FUNCTION_BLOCK "Auto_Test"   // FB1, SCL
{ S7_Optimized_Access := 'TRUE' }
VERSION : 0.1
// stored: AutoNumber true, IsIECCheckEnabled false, IsRetainMemResEnabled false, MemoryReserve 100, SetENOAutomatically false, UDAEnableTagReadback false
   VAR_INPUT
      Sys_No : UInt;
      Automatic : Bool;
      Manual : Bool;
      Level : UInt;
      Error : Bool;
      Start : Bool;
      Pause : Bool;
      Stop : Bool;
      "Pallet Type" : Char;
      "Tower 1 Pallet Alignment" : Char;
      "Tower 2 Pallet Alignment" : Char;
      "Extractor Pallet Alignment" : Char;
      Pallet_Allignment : Char;
      Tower : UInt;
      Transfer_From_To : Byte;
      "From level" : Byte;
      "To level" : Byte;
      "Testing Time" : UInt;
      "Numer of cycles" : Byte;
   END_VAR
   VAR_OUTPUT
      Running : Bool;
      Time_Runnng : Time;
      Start_Time { ExternalAccessible := 'False'; ExternalVisible := 'False'; ExternalWritable := 'False'} : String;
      Stop_Time { ExternalAccessible := 'False'; ExternalVisible := 'False'; ExternalWritable := 'False'} : String;
      Duration : Time;
   END_VAR
   VAR_IN_OUT
      "Order Table_1" : "OrderTable_UDT";
      Step_Table_0 : "OrderTable_UDT";
      System_OrderSent : Bool;
      Total_Duration : Time;
   END_VAR
   VAR
      State : Int;
      R_Start { S7_SetPoint := 'True'} : R_TRIG;
      T_Delay { S7_SetPoint := 'True'} : TON_TIME;
      Time_Delay : Time := T#0ms;
      Send_VTD_Order : Bool;
      Send_CNV_Order : Bool;
      R_TRIG_Instance { S7_SetPoint := 'True'} : R_TRIG;
      T_Running { S7_SetPoint := 'True'} : TON_TIME;
      F_TRIG { S7_SetPoint := 'True'} : F_TRIG;
      R_TRIG { S7_SetPoint := 'True'} : R_TRIG;
      Error_Code : Int;
      test : Bool;
      N_Cycles : UInt;
      Testing_Time : Time;
      R_Manual_Mode { S7_SetPoint := 'True'} : R_TRIG;
   END_VAR
   VAR_TEMP
      Busy : Bool;
   END_VAR
   VAR CONSTANT
      VTD_DEVICE : String := 'VTD';
      PALLET_INOUT_DEVICE : String := 'Pallet In Out';
      SHUTTLE_INOUT_DEVICE : String := 'Shuttle In Out';
      RUNNING_STATUS : String := 'Running';
      COMPLETED_STATUS : String := 'Completed';
   END_VAR
BEGIN
   #R_Start(CLK:=#Start);

   IF #Stop THEN
       #State := 0;
   END_IF;

   IF #Error THEN
       #State := 400;
   END_IF;

   #R_Manual_Mode(CLK:=#Automatic AND NOT #Error AND #Manual AND NOT #Running);

   IF #R_Manual_Mode.Q THEN
       #State := 500;
   ELSIF #Automatic AND NOT #Error AND NOT #Manual AND #State = 500 THEN
       #State := 0;
   END_IF;

   IF #State > 10 AND #State < 400 THEN
       #Running := TRUE;
   END_IF;

   //Time running
   #R_TRIG(CLK:=#Running);
   IF #R_TRIG.Q THEN
       #Start_Time := "Time".CurrentLocalTime;
       #Stop_Time := '';
   END_IF;
   #F_TRIG(CLK:=#Running);
   IF #F_TRIG.Q THEN
       #Duration := #T_Running.ET;
       #Total_Duration := #Duration + #Total_Duration;
       #Stop_Time := "Time".CurrentLocalTime;
   END_IF;
   #T_Running(IN:=#Running AND NOT #Pause,
                         PT:=t#24h);

   #Time_Runnng := #T_Running.ET;

   #Testing_Time := UINT_TO_TIME(#"Testing Time") * 60000;

   #Error_Code := WRIT_DBL(REQ := #test, SRCBLK := "Auto_Test_DB",BUSY=>#Busy, DSTBLK => "Auto_Test_DB");

   CASE #State OF
       0://Initialization
           #Running := false;
           #State := #State + 10;

       10://Idle
           IF #R_Start.Q AND #Automatic AND NOT #Error AND #"Pallet Type" <> '' AND #"From level" > 0 AND #"To level" > 0  THEN
               #N_Cycles := 0;
               #State := #State + 10;
           END_IF;

       20: //VTD TO START LEVEL
           IF "Control_DB".VTD_Sys[#Sys_No].Current_Level <> #"From level" THEN
               "VTD_Order_FC"(i_Sys := #Sys_No,
                              Level := #"From level",
                              StepTable_0 := #Step_Table_0);
               #R_TRIG_Instance(CLK := TRUE,
                                Q => #System_OrderSent);
               #T_Delay(IN := TRUE,
                        PT := #Time_Delay);
               IF #"Order Table_1".Status = #RUNNING_STATUS AND #T_Delay.Q THEN
                   #R_TRIG_Instance(CLK := FALSE,
                                    Q => #System_OrderSent);
                   #T_Delay(IN := FALSE,
                            PT := T#0ms);
                   #State := #State + 10;
               END_IF;
           ELSE
               #State := #State + 20;
           END_IF;

       30: //ACK VTD
           //Wait to complete and send ack
           IF #"Order Table_1".Status = #COMPLETED_STATUS AND NOT #Pause THEN
               "Control_DB".WCS_OPC_Control[#Sys_No].Movement_Request_Complete_Ack := TRUE;
               #State := #State + 10;
           END_IF;

       40: //CNV1
           "CNV_Order_FC"(i_Sys := #Sys_No,
                          Level := "Control_DB".VTD_Sys[#Sys_No].Current_Level,
                          Tower := 1,
                          Transfer_From_To := 2,
                          Pallet_Type := #"Pallet Type",
                          Pallet_Allignment := #"Tower 1 Pallet Alignment",
                          Device:=#PALLET_INOUT_DEVICE,
                          Task_Type:=4,
                          StepTable_0 := #Step_Table_0);
           #System_OrderSent := TRUE;
           #State := #State + 10;

       50: //RESET ACK
           IF #"Order Table_1".Status = #RUNNING_STATUS THEN
               "Control_DB".WCS_OPC_Control[#Sys_No].Movement_Request_Complete_Ack := FALSE;
               #R_TRIG_Instance(CLK := FALSE,
                                Q => #System_OrderSent);
               #State := #State + 10;
           END_IF;

       60: //ACK CNV1
           //Wait to complete and send ack
           IF #"Order Table_1".Status = #COMPLETED_STATUS AND NOT #Pause THEN
               "Control_DB".WCS_OPC_Control[#Sys_No].Movement_Request_Complete_Ack := TRUE;
               #State := #State + 10;
           END_IF;

       70: //ECVN TO TOWER 1
           "CNV_Order_FC"(i_Sys := #Sys_No,
                          Level := "Control_DB".VTD_Sys[#Sys_No].Current_Level,
                          Tower := 1,
                          Transfer_From_To := 1,
                          Pallet_Type := #"Pallet Type",
                          Pallet_Allignment := #"Extractor Pallet Alignment",
                          Device:=#PALLET_INOUT_DEVICE,
                          Task_Type:=4,
                          StepTable_0 := #Step_Table_0);
           #System_OrderSent := TRUE;
           #State := #State + 10;

       80: //RESET ACK
           IF #"Order Table_1".Status = #RUNNING_STATUS THEN
               "Control_DB".WCS_OPC_Control[#Sys_No].Movement_Request_Complete_Ack := FALSE;
               #State := #State + 10;
           END_IF;

       90: //ACK ECVN
           //Wait to complete and send ack
           IF #"Order Table_1".Status = #COMPLETED_STATUS AND NOT #Pause THEN
               "Control_DB".WCS_OPC_Control[#Sys_No].Movement_Request_Complete_Ack := TRUE;
               #State := #State + 10;
           END_IF;

       100: //VTD FROM START LEVEL TO FINAL LEVEL
           IF "Control_DB".VTD_Sys[#Sys_No].Current_Level < #"To level" THEN
               "VTD_Order_FC"(i_Sys := #Sys_No,
                              Level := "Control_DB".VTD_Sys[#Sys_No].Current_Level + 1,
                              StepTable_0 := #Step_Table_0);
               #System_OrderSent := TRUE;
               #State := #State + 10;
           ELSE
               #State := 130;
           END_IF;

       110: //RESET ACK
           IF #"Order Table_1".Status = #RUNNING_STATUS THEN
               "Control_DB".WCS_OPC_Control[#Sys_No].Movement_Request_Complete_Ack := FALSE;
               #State := #State + 10;
           END_IF;


       120: //ACK VTD
           //Wait to complete and send ack
           IF #"Order Table_1".Status = #COMPLETED_STATUS AND NOT #Pause THEN
               "Control_DB".WCS_OPC_Control[#Sys_No].Movement_Request_Complete_Ack := TRUE;
               #State := 40;
           END_IF;

       130: //VTD TO START LEVEL---------------------------------------------------------------------------------------------------
           "VTD_Order_FC"(i_Sys := #Sys_No,
                          Level := #"From level",
                          StepTable_0 := #Step_Table_0);
           #System_OrderSent := TRUE;
           #State := #State + 10;

       140: //RESET ACK
           IF #"Order Table_1".Status = #RUNNING_STATUS THEN
               "Control_DB".WCS_OPC_Control[#Sys_No].Movement_Request_Complete_Ack := FALSE;
               #State := #State + 10;
           END_IF;

       150: //ACK VTD START LEVEL
           //Wait to complete and send ack
           IF #Sys_No <= 3 THEN
               IF #"Order Table_1".Status = #COMPLETED_STATUS AND NOT #Pause THEN
                   "Control_DB".WCS_OPC_Control[#Sys_No].Movement_Request_Complete_Ack := TRUE;
                   #State := #State + 10;
               END_IF;
           ELSE
               IF #"Order Table_1".Status = #COMPLETED_STATUS AND NOT #Pause THEN
                   "Control_DB".WCS_OPC_Control[#Sys_No].Movement_Request_Complete_Ack := TRUE;
                   #State := 40; //TEST JUST CONV 1 FOR SYSTEM 4 AND 5
               END_IF;
           END_IF;

       160: //CNV2
           "CNV_Order_FC"(i_Sys := #Sys_No,
                          Level := "Control_DB".VTD_Sys[#Sys_No].Current_Level,
                          Tower := 2,
                          Transfer_From_To := 2,
                          Pallet_Type := #"Pallet Type",
                          Pallet_Allignment := #"Tower 2 Pallet Alignment",
                          Device:=#PALLET_INOUT_DEVICE,
                          Task_Type:=4,
                          StepTable_0 := #Step_Table_0);
           #System_OrderSent := TRUE;
           #State := #State + 10;

       170: //RESET ACK
           IF #"Order Table_1".Status = #RUNNING_STATUS THEN
               "Control_DB".WCS_OPC_Control[#Sys_No].Movement_Request_Complete_Ack := FALSE;
               #State := #State + 10;
           END_IF;

       180: //ACK CNV2
           //Wait to complete and send ack
           IF #"Order Table_1".Status = #COMPLETED_STATUS AND NOT #Pause THEN
               "Control_DB".WCS_OPC_Control[#Sys_No].Movement_Request_Complete_Ack := TRUE;
               #State := #State + 10;
           END_IF;

       190: //ECVN TO TOWER 2
           "CNV_Order_FC"(i_Sys := #Sys_No,
                          Level := "Control_DB".VTD_Sys[#Sys_No].Current_Level,
                          Tower := 2,
                          Transfer_From_To := 1,
                          Pallet_Type := #"Pallet Type",
                          Pallet_Allignment := #"Extractor Pallet Alignment",
                          Device:=#PALLET_INOUT_DEVICE,
                          Task_Type:=4,
                          StepTable_0 := #Step_Table_0);
           #System_OrderSent := TRUE;
           #State := #State + 10;

       200: //RESET ACK
           IF #"Order Table_1".Status = #RUNNING_STATUS THEN
               "Control_DB".WCS_OPC_Control[#Sys_No].Movement_Request_Complete_Ack := FALSE;
               #State := #State + 10;
           END_IF;

       210: //ACK ECVN TO TOWER 2
           //Wait to complete and send ack
           IF #"Order Table_1".Status = #COMPLETED_STATUS AND NOT #Pause THEN
               "Control_DB".WCS_OPC_Control[#Sys_No].Movement_Request_Complete_Ack := TRUE;
               #State := #State + 10;
           END_IF;

       220: //VTD 
           IF "Control_DB".VTD_Sys[#Sys_No].Current_Level < #"To level" THEN
               "VTD_Order_FC"(i_Sys := #Sys_No,
                              Level := "Control_DB".VTD_Sys[#Sys_No].Current_Level + 1,
                              StepTable_0 := #Step_Table_0);
               #System_OrderSent := TRUE;
               #State := #State + 10;
           ELSIF (
               (#"Numer of cycles" = 0 OR #N_Cycles < #"Numer of cycles")
               AND
               (#Testing_Time = T#0M OR #Time_Runnng < #Testing_Time)
               ) THEN
               #State := 250;//CONTINUE
           ELSE
               #State := 260;//FINISH
           END_IF;

       230: //RESET ACK
           IF #"Order Table_1".Status = #RUNNING_STATUS THEN
               "Control_DB".WCS_OPC_Control[#Sys_No].Movement_Request_Complete_Ack := FALSE;
               #State := #State + 10;
           END_IF;

       240: //ACK VTD
           //Wait to complete and send ack
           IF #"Order Table_1".Status = #COMPLETED_STATUS AND NOT #Pause THEN
               "Control_DB".WCS_OPC_Control[#Sys_No].Movement_Request_Complete_Ack := TRUE;
               #State := 160;
           END_IF;

       250: //ACK VTD AND START ANOTHER CYCLE
           //Wait to complete and send ack
           IF #"Order Table_1".Status = #COMPLETED_STATUS AND NOT #Pause THEN
               "Control_DB".WCS_OPC_Control[#Sys_No].Movement_Request_Complete_Ack := TRUE;
               #N_Cycles := #N_Cycles + 1;
               #State := 20;
           END_IF;

       260: //ACK VTD AND FINISH
           //Wait to complete and send ack
           IF #"Order Table_1".Status = #COMPLETED_STATUS AND NOT #Pause THEN
               "Control_DB".WCS_OPC_Control[#Sys_No].Movement_Request_Complete_Ack := TRUE;
               #State := 0;
           END_IF;

       400: //ERROR
           #Running := false;
           IF "Reset_All" OR
               ("Screen_DB_1".Reset_All[1] AND
                ("HMI_Box_Connected_1" = 1) OR ("HMI_Box_Connected_1" = 2) OR ("HMI_Box_Connected_1" = 3) OR ("HMI_Box_Connected_1" = 4) OR ("HMI_Box_Connected_1" = 5) OR
                ("HMI_Box_Connected_1" = 11 AND "KEY REMOTE/LOCAL L1 - CH1(1)") OR
                ("HMI_Box_Connected_1" = 12 AND "KEY REMOTE/LOCAL L2 - CH1(1)") OR
                ("HMI_Box_Connected_1" = 13 AND "KEY REMOTE/LOCAL L3 - CH1(1)") OR
                ("HMI_Box_Connected_1" = 14 AND "KEY REMOTE/LOCAL L4 - CH1(1)") OR
                ("HMI_Box_Connected_1" = 15 AND "KEY REMOTE/LOCAL L5 - CH1(1)") OR
                ("HMI_Box_Connected_1" = 16 AND "KEY REMOTE/LOCAL L6 - CH1(1)") OR
                ("HMI_Box_Connected_1" = 17 AND "KEY REMOTE/LOCAL L7 - CH1(1)") OR
                ("HMI_Box_Connected_1" = 18 AND "KEY REMOTE/LOCAL L8 - CH1(1)") OR
                ("HMI_Box_Connected_1" = 21 AND "KEY REMOTE/LOCAL L1 - CH1(2)") OR
                ("HMI_Box_Connected_1" = 22 AND "KEY REMOTE/LOCAL L2 - CH1(2)") OR
                ("HMI_Box_Connected_1" = 23 AND "KEY REMOTE/LOCAL L3 - CH1(2)") OR
                ("HMI_Box_Connected_1" = 24 AND "KEY REMOTE/LOCAL L4 - CH1(2)") OR
                ("HMI_Box_Connected_1" = 25 AND "KEY REMOTE/LOCAL L5 - CH1(2)") OR
                ("HMI_Box_Connected_1" = 26 AND "KEY REMOTE/LOCAL L6 - CH1(2)") OR
                ("HMI_Box_Connected_1" = 27 AND "KEY REMOTE/LOCAL L7 - CH1(2)") OR
                ("HMI_Box_Connected_1" = 28 AND "KEY REMOTE/LOCAL L8 - CH1(2)") OR
                ("HMI_Box_Connected_1" = 31 AND "KEY REMOTE/LOCAL L1 - CH1(3)") OR
                ("HMI_Box_Connected_1" = 32 AND "KEY REMOTE/LOCAL L2 - CH1(3)") OR
                ("HMI_Box_Connected_1" = 33 AND "KEY REMOTE/LOCAL L3 - CH1(3)") OR
                ("HMI_Box_Connected_1" = 34 AND "KEY REMOTE/LOCAL L4 - CH1(3)") OR
                ("HMI_Box_Connected_1" = 35 AND "KEY REMOTE/LOCAL L5 - CH1(3)") OR
                ("HMI_Box_Connected_1" = 36 AND "KEY REMOTE/LOCAL L6 - CH1(3)") OR
                ("HMI_Box_Connected_1" = 37 AND "KEY REMOTE/LOCAL L7 - CH1(3)") OR
                ("HMI_Box_Connected_1" = 38 AND "KEY REMOTE/LOCAL L8 - CH1(3)") OR
                ("HMI_Box_Connected_1" = 41 AND "KEY REMOTE/LOCAL L1 - CH1(4)") OR
                ("HMI_Box_Connected_1" = 42 AND "KEY REMOTE/LOCAL L2 - CH1(4)") OR
                ("HMI_Box_Connected_1" = 43 AND "KEY REMOTE/LOCAL L3 - CH1(4)") OR
                ("HMI_Box_Connected_1" = 44 AND "KEY REMOTE/LOCAL L4 - CH1(4)") OR
                ("HMI_Box_Connected_1" = 45 AND "KEY REMOTE/LOCAL L5 - CH1(4)") OR
                ("HMI_Box_Connected_1" = 46 AND "KEY REMOTE/LOCAL L6 - CH1(4)") OR
                ("HMI_Box_Connected_1" = 47 AND "KEY REMOTE/LOCAL L7 - CH1(4)") OR
                ("HMI_Box_Connected_1" = 48 AND "KEY REMOTE/LOCAL L8 - CH1(4)") OR
                ("HMI_Box_Connected_1" = 51 AND "KEY REMOTE/LOCAL L1 - CH1(5)") OR
                ("HMI_Box_Connected_1" = 52 AND "KEY REMOTE/LOCAL L2 - CH1(5)") OR
                ("HMI_Box_Connected_1" = 53 AND "KEY REMOTE/LOCAL L3 - CH1(5)") OR
                ("HMI_Box_Connected_1" = 54 AND "KEY REMOTE/LOCAL L4 - CH1(5)") OR
                ("HMI_Box_Connected_1" = 55 AND "KEY REMOTE/LOCAL L5 - CH1(5)") OR
                ("HMI_Box_Connected_1" = 56 AND "KEY REMOTE/LOCAL L6 - CH1(5)") OR
                ("HMI_Box_Connected_1" = 57 AND "KEY REMOTE/LOCAL L7 - CH1(5)") OR
                ("HMI_Box_Connected_1" = 58 AND "KEY REMOTE/LOCAL L8 - CH1(5)"))
           THEN
               #State := 0;
           END_IF;

       500://MANUAL ORDER
           #Running := false;
           IF #Send_VTD_Order THEN
               "VTD_Order_FC"(i_Sys := #Sys_No,
                              Level := #Level,
                              StepTable_0 := #Step_Table_0);
               #System_OrderSent := TRUE;
               #Running := TRUE;
               #Send_VTD_Order := FALSE;
           END_IF;

           IF #Send_CNV_Order THEN
               "CNV_Order_FC"(i_Sys := #Sys_No,
                              Level := "Control_DB".VTD_Sys[#Sys_No].Current_Level,
                              Tower := #Tower,
                              Transfer_From_To := #Transfer_From_To,
                              Pallet_Type := #"Pallet Type",
                              Pallet_Allignment := #Pallet_Allignment,
                              Device:=#PALLET_INOUT_DEVICE,
                              Task_Type:=4,
                              StepTable_0 := #Step_Table_0);
               #System_OrderSent := TRUE;
               #Running := TRUE;
               #Send_CNV_Order := FALSE;
           END_IF;

           IF #"Order Table_1".Status = #RUNNING_STATUS THEN
               #State := #State + 10;
           END_IF;

       510: //RESET ACK
           IF #"Order Table_1".Status = #RUNNING_STATUS THEN
               "Control_DB".WCS_OPC_Control[#Sys_No].Movement_Request_Complete_Ack := FALSE;
               #State := #State + 10;
           END_IF;

       520: //ACK VTD
           //Wait to complete and send ack
           IF #"Order Table_1".Status = #COMPLETED_STATUS THEN
               "Control_DB".WCS_OPC_Control[#Sys_No].Movement_Request_Complete_Ack := TRUE;
               #State := 500;
           END_IF;
   END_CASE;
END_FUNCTION_BLOCK

FUNCTION_BLOCK "Auto_Test_1"   // FB3, SCL
{ S7_Optimized_Access := 'TRUE' }
VERSION : 0.1
// stored: AutoNumber true, IsIECCheckEnabled false, IsRetainMemResEnabled false, MemoryReserve 100, SetENOAutomatically false, UDAEnableTagReadback false
   VAR_INPUT
      Sys_No : UInt;
      Automatic : Bool;
      Manual : Bool;
      Level : UInt;
      Error : Bool;
      Start : Bool;
      Pause : Bool;
      Stop : Bool;
      "Pallet Type" : Char;
      "Tower 1 Pallet Alignment" : Char;
      "Tower 2 Pallet Alignment" : Char;
      "Extractor Pallet Alignment" : Char;
      Pallet_Allignment : Char;
      Tower : UInt;
      Transfer_From_To : Byte;
      "From level" : Byte;
      "To level" : Byte;
      "Testing Time" : UInt;
      "Numer of cycles" : Byte;
   END_VAR
   VAR_OUTPUT
      Running : Bool;
      Time_Runnng : Time;
      Start_Time { ExternalAccessible := 'False'; ExternalVisible := 'False'; ExternalWritable := 'False'} : String;
      Stop_Time { ExternalAccessible := 'False'; ExternalVisible := 'False'; ExternalWritable := 'False'} : String;
      Duration : Time;
   END_VAR
   VAR_IN_OUT
      "Order Table_1" : "OrderTable_UDT";
      Step_Table_0 : "OrderTable_UDT";
      System_OrderSent : Bool;
      Total_Duration : Time;
   END_VAR
   VAR
      State : Int;
      R_Start { S7_SetPoint := 'True'} : R_TRIG;
      T_Delay { S7_SetPoint := 'True'} : TON_TIME;
      Time_Delay : Time := T#0ms;
      Send_VTD_Order : Bool;
      Send_CNV_Order : Bool;
      R_TRIG_Instance { S7_SetPoint := 'True'} : R_TRIG;
      T_Running { S7_SetPoint := 'True'} : TON_TIME;
      F_TRIG { S7_SetPoint := 'True'} : F_TRIG;
      R_TRIG { S7_SetPoint := 'True'} : R_TRIG;
      Error_Code : Int;
      test : Bool;
      N_Cycles : UInt;
      Testing_Time : Time;
      R_Manual_Mode { S7_SetPoint := 'True'} : R_TRIG;
   END_VAR
   VAR_TEMP
      Busy : Bool;
   END_VAR
   VAR CONSTANT
      VTD_DEVICE : String := 'VTD';
      PALLET_INOUT_DEVICE : String := 'Pallet In Out';
      SHUTTLE_INOUT_DEVICE : String := 'Shuttle In Out';
      RUNNING_STATUS : String := 'Running';
      COMPLETED_STATUS : String := 'Completed';
   END_VAR
BEGIN
   #R_Start(CLK:=#Start);

   IF #Stop THEN
       #State := 0;
   END_IF;

   IF #Error THEN
       #State := 400;
   END_IF;

   #R_Manual_Mode(CLK:=#Automatic AND NOT #Error AND #Manual AND NOT #Running);

   IF #R_Manual_Mode.Q THEN
       #State := 500;
   ELSIF #Automatic AND NOT #Error AND NOT #Manual AND #State = 500 THEN
       #State := 0;
   END_IF;

   IF #State > 10 AND #State < 400 THEN
       #Running := TRUE;
   END_IF;

   //Time running
   #R_TRIG(CLK:=#Running);
   IF #R_TRIG.Q THEN
       #Start_Time := "Time".CurrentLocalTime;
       #Stop_Time := '';
   END_IF;
   #F_TRIG(CLK:=#Running);
   IF #F_TRIG.Q THEN
       #Duration := #T_Running.ET;
       #Total_Duration := #Duration + #Total_Duration;
       #Stop_Time := "Time".CurrentLocalTime;
   END_IF;
   #T_Running(IN:=#Running AND NOT #Pause,
                         PT:=t#24h);

   #Time_Runnng := #T_Running.ET;

   #Testing_Time := UINT_TO_TIME(#"Testing Time") * 60000;

   #Error_Code := WRIT_DBL(REQ := #test, SRCBLK := "Auto_Test_DB",BUSY=>#Busy, DSTBLK => "Auto_Test_DB");

   CASE #State OF
       0://Initialization
           #Running := false;
           #State := #State + 10;

       10://Idle
           IF #R_Start.Q AND #Automatic AND NOT #Error AND #"Pallet Type" <> '' AND #"From level" > 0 AND #"To level" > 0  THEN
               #N_Cycles := 0;
               #State := #State + 10;
           END_IF;

       20: //VTD TO START LEVEL
           IF "Control_DB".VTD_Sys[#Sys_No].Current_Level <> #"From level" THEN
               "VTD_Order_FC"(i_Sys := #Sys_No,
                              Level := #"From level",
                              StepTable_0 := #Step_Table_0);
               #R_TRIG_Instance(CLK := TRUE,
                                Q => #System_OrderSent);
               #T_Delay(IN := TRUE,
                        PT := #Time_Delay);
               IF #"Order Table_1".Status = #RUNNING_STATUS AND #T_Delay.Q THEN
                   #R_TRIG_Instance(CLK := FALSE,
                                    Q => #System_OrderSent);
                   #T_Delay(IN := FALSE,
                            PT := T#0ms);
                   #State := #State + 10;
               END_IF;
           ELSE
               #State := #State + 20;
           END_IF;

       30: //ACK VTD
           //Wait to complete and send ack
           IF #"Order Table_1".Status = #COMPLETED_STATUS AND NOT #Pause THEN
               "Control_DB".WCS_OPC_Control[#Sys_No].Movement_Request_Complete_Ack := TRUE;
               #State := #State + 10;
           END_IF;

       40: //CNV1
           "CNV_Order_FC"(i_Sys := #Sys_No,
                          Level := "Control_DB".VTD_Sys[#Sys_No].Current_Level,
                          Tower := 1,
                          Transfer_From_To := 2,
                          Pallet_Type := #"Pallet Type",
                          Pallet_Allignment := #"Tower 1 Pallet Alignment",
                          Device:=#PALLET_INOUT_DEVICE,
                          Task_Type:=4,
                          StepTable_0 := #Step_Table_0);
           #System_OrderSent := TRUE;
           #State := #State + 10;

       50: //RESET ACK
           IF #"Order Table_1".Status = #RUNNING_STATUS THEN
               "Control_DB".WCS_OPC_Control[#Sys_No].Movement_Request_Complete_Ack := FALSE;
               #R_TRIG_Instance(CLK := FALSE,
                                Q => #System_OrderSent);
               #State := #State + 10;
           END_IF;

       60: //ACK CNV1
           //Wait to complete and send ack
           IF #"Order Table_1".Status = #COMPLETED_STATUS AND NOT #Pause THEN
               "Control_DB".WCS_OPC_Control[#Sys_No].Movement_Request_Complete_Ack := TRUE;
               #State := #State + 10;
           END_IF;

       70: //ECVN TO TOWER 1
           "CNV_Order_FC"(i_Sys := #Sys_No,
                          Level := "Control_DB".VTD_Sys[#Sys_No].Current_Level,
                          Tower := 1,
                          Transfer_From_To := 1,
                          Pallet_Type := #"Pallet Type",
                          Pallet_Allignment := #"Extractor Pallet Alignment",
                          Device:=#PALLET_INOUT_DEVICE,
                          Task_Type:=4,
                          StepTable_0 := #Step_Table_0);
           #System_OrderSent := TRUE;
           #State := #State + 10;

       80: //RESET ACK
           IF #"Order Table_1".Status = #RUNNING_STATUS THEN
               "Control_DB".WCS_OPC_Control[#Sys_No].Movement_Request_Complete_Ack := FALSE;
               #State := #State + 10;
           END_IF;

       90: //ACK ECVN
           //Wait to complete and send ack
           IF #"Order Table_1".Status = #COMPLETED_STATUS AND NOT #Pause THEN
               "Control_DB".WCS_OPC_Control[#Sys_No].Movement_Request_Complete_Ack := TRUE;
               #State := #State + 10;
           END_IF;

       100: //VTD FROM START LEVEL TO FINAL LEVEL
           IF "Control_DB".VTD_Sys[#Sys_No].Current_Level < #"To level" THEN
               "VTD_Order_FC"(i_Sys := #Sys_No,
                              Level := "Control_DB".VTD_Sys[#Sys_No].Current_Level + 1,
                              StepTable_0 := #Step_Table_0);
               #System_OrderSent := TRUE;
               #State := #State + 10;
           ELSIF (
               (#"Numer of cycles" = 0 OR #N_Cycles < #"Numer of cycles")
               AND
               (#Testing_Time = T#0M OR #Time_Runnng < #Testing_Time)
               ) THEN
               #State := 250;//CONTINUE
           ELSE
               #State := 260;//FINISH
           END_IF;

       110: //RESET ACK
           IF #"Order Table_1".Status = #RUNNING_STATUS THEN
               "Control_DB".WCS_OPC_Control[#Sys_No].Movement_Request_Complete_Ack := FALSE;
               #State := #State + 10;
           END_IF;


       120: //ACK VTD
           //Wait to complete and send ack
           IF #"Order Table_1".Status = #COMPLETED_STATUS AND NOT #Pause THEN
               "Control_DB".WCS_OPC_Control[#Sys_No].Movement_Request_Complete_Ack := TRUE;
               #State := 40;
           END_IF;

       250: //ACK VTD AND START ANOTHER CYCLE
           //Wait to complete and send ack
           IF #"Order Table_1".Status = #COMPLETED_STATUS AND NOT #Pause THEN
               "Control_DB".WCS_OPC_Control[#Sys_No].Movement_Request_Complete_Ack := TRUE;
               #N_Cycles := #N_Cycles + 1;
               #State := 20;
           END_IF;

       260: //ACK VTD AND FINISH
           //Wait to complete and send ack
           IF #"Order Table_1".Status = #COMPLETED_STATUS AND NOT #Pause THEN
               "Control_DB".WCS_OPC_Control[#Sys_No].Movement_Request_Complete_Ack := TRUE;
               #State := 0;
           END_IF;

       400: //ERROR
           #Running := false;
           IF "Reset_All" OR
               ("Screen_DB_1".Reset_All[1] AND
                ("HMI_Box_Connected_1" = 1) OR ("HMI_Box_Connected_1" = 2) OR ("HMI_Box_Connected_1" = 3) OR ("HMI_Box_Connected_1" = 4) OR ("HMI_Box_Connected_1" = 5) OR
                ("HMI_Box_Connected_1" = 11 AND "KEY REMOTE/LOCAL L1 - CH1(1)") OR
                ("HMI_Box_Connected_1" = 12 AND "KEY REMOTE/LOCAL L2 - CH1(1)") OR
                ("HMI_Box_Connected_1" = 13 AND "KEY REMOTE/LOCAL L3 - CH1(1)") OR
                ("HMI_Box_Connected_1" = 14 AND "KEY REMOTE/LOCAL L4 - CH1(1)") OR
                ("HMI_Box_Connected_1" = 15 AND "KEY REMOTE/LOCAL L5 - CH1(1)") OR
                ("HMI_Box_Connected_1" = 16 AND "KEY REMOTE/LOCAL L6 - CH1(1)") OR
                ("HMI_Box_Connected_1" = 17 AND "KEY REMOTE/LOCAL L7 - CH1(1)") OR
                ("HMI_Box_Connected_1" = 18 AND "KEY REMOTE/LOCAL L8 - CH1(1)") OR
                ("HMI_Box_Connected_1" = 21 AND "KEY REMOTE/LOCAL L1 - CH1(2)") OR
                ("HMI_Box_Connected_1" = 22 AND "KEY REMOTE/LOCAL L2 - CH1(2)") OR
                ("HMI_Box_Connected_1" = 23 AND "KEY REMOTE/LOCAL L3 - CH1(2)") OR
                ("HMI_Box_Connected_1" = 24 AND "KEY REMOTE/LOCAL L4 - CH1(2)") OR
                ("HMI_Box_Connected_1" = 25 AND "KEY REMOTE/LOCAL L5 - CH1(2)") OR
                ("HMI_Box_Connected_1" = 26 AND "KEY REMOTE/LOCAL L6 - CH1(2)") OR
                ("HMI_Box_Connected_1" = 27 AND "KEY REMOTE/LOCAL L7 - CH1(2)") OR
                ("HMI_Box_Connected_1" = 28 AND "KEY REMOTE/LOCAL L8 - CH1(2)") OR
                ("HMI_Box_Connected_1" = 31 AND "KEY REMOTE/LOCAL L1 - CH1(3)") OR
                ("HMI_Box_Connected_1" = 32 AND "KEY REMOTE/LOCAL L2 - CH1(3)") OR
                ("HMI_Box_Connected_1" = 33 AND "KEY REMOTE/LOCAL L3 - CH1(3)") OR
                ("HMI_Box_Connected_1" = 34 AND "KEY REMOTE/LOCAL L4 - CH1(3)") OR
                ("HMI_Box_Connected_1" = 35 AND "KEY REMOTE/LOCAL L5 - CH1(3)") OR
                ("HMI_Box_Connected_1" = 36 AND "KEY REMOTE/LOCAL L6 - CH1(3)") OR
                ("HMI_Box_Connected_1" = 37 AND "KEY REMOTE/LOCAL L7 - CH1(3)") OR
                ("HMI_Box_Connected_1" = 38 AND "KEY REMOTE/LOCAL L8 - CH1(3)") OR
                ("HMI_Box_Connected_1" = 41 AND "KEY REMOTE/LOCAL L1 - CH1(4)") OR
                ("HMI_Box_Connected_1" = 42 AND "KEY REMOTE/LOCAL L2 - CH1(4)") OR
                ("HMI_Box_Connected_1" = 43 AND "KEY REMOTE/LOCAL L3 - CH1(4)") OR
                ("HMI_Box_Connected_1" = 44 AND "KEY REMOTE/LOCAL L4 - CH1(4)") OR
                ("HMI_Box_Connected_1" = 45 AND "KEY REMOTE/LOCAL L5 - CH1(4)") OR
                ("HMI_Box_Connected_1" = 46 AND "KEY REMOTE/LOCAL L6 - CH1(4)") OR
                ("HMI_Box_Connected_1" = 47 AND "KEY REMOTE/LOCAL L7 - CH1(4)") OR
                ("HMI_Box_Connected_1" = 48 AND "KEY REMOTE/LOCAL L8 - CH1(4)") OR
                ("HMI_Box_Connected_1" = 51 AND "KEY REMOTE/LOCAL L1 - CH1(5)") OR
                ("HMI_Box_Connected_1" = 52 AND "KEY REMOTE/LOCAL L2 - CH1(5)") OR
                ("HMI_Box_Connected_1" = 53 AND "KEY REMOTE/LOCAL L3 - CH1(5)") OR
                ("HMI_Box_Connected_1" = 54 AND "KEY REMOTE/LOCAL L4 - CH1(5)") OR
                ("HMI_Box_Connected_1" = 55 AND "KEY REMOTE/LOCAL L5 - CH1(5)") OR
                ("HMI_Box_Connected_1" = 56 AND "KEY REMOTE/LOCAL L6 - CH1(5)") OR
                ("HMI_Box_Connected_1" = 57 AND "KEY REMOTE/LOCAL L7 - CH1(5)") OR
                ("HMI_Box_Connected_1" = 58 AND "KEY REMOTE/LOCAL L8 - CH1(5)"))
           THEN
               #State := 0;
           END_IF;

       500://MANUAL ORDER
           #Running := false;
           IF #Send_VTD_Order THEN
               "VTD_Order_FC"(i_Sys := #Sys_No,
                              Level := #Level,
                              StepTable_0 := #Step_Table_0);
               #System_OrderSent := TRUE;
               #Running := TRUE;
               #Send_VTD_Order := FALSE;
           END_IF;

           IF #Send_CNV_Order THEN
               "CNV_Order_FC"(i_Sys := #Sys_No,
                              Level := "Control_DB".VTD_Sys[#Sys_No].Current_Level,
                              Tower := #Tower,
                              Transfer_From_To := #Transfer_From_To,
                              Pallet_Type := #"Pallet Type",
                              Pallet_Allignment := #Pallet_Allignment,
                              Device:=#PALLET_INOUT_DEVICE,
                              Task_Type:=4,
                              StepTable_0 := #Step_Table_0);
               #System_OrderSent := TRUE;
               #Running := TRUE;
               #Send_CNV_Order := FALSE;
           END_IF;

           IF #"Order Table_1".Status = #RUNNING_STATUS THEN
               #State := #State + 10;
           END_IF;

       510: //RESET ACK
           IF #"Order Table_1".Status = #RUNNING_STATUS THEN
               "Control_DB".WCS_OPC_Control[#Sys_No].Movement_Request_Complete_Ack := FALSE;
               #State := #State + 10;
           END_IF;

       520: //ACK VTD
           //Wait to complete and send ack
           IF #"Order Table_1".Status = #COMPLETED_STATUS THEN
               "Control_DB".WCS_OPC_Control[#Sys_No].Movement_Request_Complete_Ack := TRUE;
               #State := 500;
           END_IF;
   END_CASE;
END_FUNCTION_BLOCK

FUNCTION "Conveyors_Transfer" : Void   // FC24, SCL
{ S7_Optimized_Access := 'TRUE' }
VERSION : 0.1
// stored: AutoNumber true, IsIECCheckEnabled false, SetENOAutomatically false, UDAEnableTagReadback false
   VAR_TEMP
      i_Lev : UInt;
      i_Sys : UInt;
      Concat1 : String;
      Concat2 : String;
      ID : DInt;
      StrLev : String;
      StrSys : String;
      Level : UInt;
   END_VAR
BEGIN
   FOR #i_Sys := 1 TO 5 DO
       #StrSys := UINT_TO_STRING(#i_Sys);
       // Remove "+"
       IF #StrSys[1] = '+' THEN
           #StrSys := RIGHT(IN := #StrSys, L := LEN(#StrSys) - 1);
       END_IF;

       REGION ID OF THE VTD CONVEYOR
           FOR #i_Lev := "Settings_DB".VTD_Sys[#i_Sys].Lowest_Level TO "Settings_DB".VTD_Sys[#i_Sys].Highest_Level DO
               IF (#i_Sys >= 1) AND (#i_Sys <= 5) THEN
                   IF "Control_DB".VTD_Sys[#i_Sys].Current_Level = #i_Lev THEN
                       #StrLev := UINT_TO_STRING(#i_Lev);

                       // Remove "+"
                       IF #StrLev[1] = '+' THEN
                           #StrLev := RIGHT(IN := #StrLev, L := LEN(#StrLev) - 1);
                       END_IF;

                       //Build ID
                       #Concat1 := CONCAT(IN1 := '120', IN2 := #StrLev);
                       #Concat2 := CONCAT(IN1 := #Concat1, IN2 := '0');
                       #ID := STRING_TO_DINT(IN := CONCAT(IN1 := #Concat2, IN2 := #StrSys));

                       "Settings_DB".ECnv_Sys[#i_Sys].ID := #ID;
                       "Settings_DB".ECnv_Sys[#i_Sys].Cnv_Level := #i_Lev;
                   END_IF;
               END_IF;
           END_FOR;
       END_REGION

           REGION READY TO RECEIVE
               //EXTRACTOR CONVEYOR
               FOR #i_Lev := "Settings_DB".VTD_Sys[#i_Sys].Lowest_Level TO "Settings_DB".VTD_Sys[#i_Sys].Highest_Level DO
                   IF "Control_DB".VTD_Sys[#i_Sys].Current_Level = #i_Lev THEN
                       #StrLev := UINT_TO_STRING(#i_Lev);

                       // Remove "+"
                       IF #StrLev[1] = '+' THEN
                           #StrLev := RIGHT(IN := #StrLev, L := LEN(#StrLev) - 1);
                       END_IF;

                       //Build ID
                       #Concat1 := CONCAT(IN1 := '120', IN2 := #StrLev);
                       #Concat2 := CONCAT(IN1 := #Concat1, IN2 := '0');
                       #ID := STRING_TO_DINT(IN := CONCAT(IN1 := #Concat2, IN2 := #StrSys));
                   END_IF;

                   IF "Settings_DB".ECnv_Sys[#i_Sys].ID = #ID AND NOT "Control_DB".ECnv_Sys[#i_Sys].Error AND NOT "Control_DB".ECnv_Sys[#i_Sys].Running
                       AND NOT "Control_DB".ECnv_Sys[#i_Sys].Cnv_Occupied AND NOT "Control_DB".ECnv_Sys[#i_Sys].Instruction.Outbound_Ready AND
                       ("Control_DB".ECnv_Sys[#i_Sys].Mode = 2 OR "Control_DB".ECnv_Sys[#i_Sys].Mode = 3) THEN
                       "Control_DB".ECnv_Sys[#i_Sys].Instruction.Inbound_Ready := TRUE;
                   ELSIF "Control_DB".ECnv_Sys[#i_Sys].Cnv_Occupied THEN  // // // // // // // // // // // // //last change
                       "Control_DB".ECnv_Sys[#i_Sys].Instruction.Inbound_Ready := FALSE;  // // // // // // // // // // // // //last change
                   END_IF;
               END_FOR;

               //BUFFER CONVEYORS
               FOR #i_Lev := "Settings_DB".VTD_Sys[#i_Sys].Lowest_Level TO "Settings_DB".VTD_Sys[#i_Sys].Highest_Level DO
                   //CNV 1
                   IF NOT "Control_DB".LCnv_Sys[#i_Sys].Cnv_Level[#i_Lev].Cnv1.Error AND
                       NOT "Control_DB".LCnv_Sys[#i_Sys].Cnv_Level[#i_Lev].Cnv1.Running AND
                       NOT "Control_DB".LCnv_Sys[#i_Sys].Cnv_Level[#i_Lev].Cnv1.Cnv_Occupied AND
                       NOT "Control_DB".LCnv_Sys[#i_Sys].Cnv_Level[#i_Lev].Cnv1.Instruction.Outbound_Ready AND
                       ("Control_DB".LCnv_Sys[#i_Sys].Cnv_Level[#i_Lev].Cnv1.Mode = 2 OR "Control_DB".LCnv_Sys[#i_Sys].Cnv_Level[#i_Lev].Cnv1.Mode = 3) AND
                       (NOT "Control_DB".ECnv_Sys[#i_Sys].Running OR "Settings_DB".LCnv_Sys[#i_Sys].Cnv_Level[#i_Lev].Cnv1.Cnv_Level <> 1)
                   THEN
                       "Control_DB".LCnv_Sys[#i_Sys].Cnv_Level[#i_Lev].Cnv1.Instruction.Inbound_Ready := TRUE;
                   ELSIF "Control_DB".LCnv_Sys[#i_Sys].Cnv_Level[#i_Lev].Cnv1.Cnv_Occupied THEN  // // // // // // // // // // // // //last change
                       "Control_DB".LCnv_Sys[#i_Sys].Cnv_Level[#i_Lev].Cnv1.Instruction.Inbound_Ready := FALSE;  // // // // // // // // // // // // //last change
                   END_IF;

                   //CNV 2
                   IF NOT "Control_DB".LCnv_Sys[#i_Sys].Cnv_Level[#i_Lev].Cnv2.Error AND
                       NOT "Control_DB".LCnv_Sys[#i_Sys].Cnv_Level[#i_Lev].Cnv2.Running AND
                       NOT "Control_DB".LCnv_Sys[#i_Sys].Cnv_Level[#i_Lev].Cnv2.Cnv_Occupied AND
                       NOT "Control_DB".LCnv_Sys[#i_Sys].Cnv_Level[#i_Lev].Cnv2.Instruction.Outbound_Ready AND
                       ("Control_DB".LCnv_Sys[#i_Sys].Cnv_Level[#i_Lev].Cnv2.Mode = 2 OR "Control_DB".LCnv_Sys[#i_Sys].Cnv_Level[#i_Lev].Cnv2.Mode = 3) THEN
                       "Control_DB".LCnv_Sys[#i_Sys].Cnv_Level[#i_Lev].Cnv2.Instruction.Inbound_Ready := TRUE;
                   ELSIF "Control_DB".LCnv_Sys[#i_Sys].Cnv_Level[#i_Lev].Cnv2.Cnv_Occupied THEN  // // // // // // // // // // // // //last change
                       "Control_DB".LCnv_Sys[#i_Sys].Cnv_Level[#i_Lev].Cnv2.Instruction.Inbound_Ready := FALSE;  // // // // // // // // // // // // //last change
                   END_IF;
               END_FOR;
           END_REGION

           REGION READY TO SEND
               //EXTRACTOR CONVEYOR
               #Level := "Settings_DB".ECnv_Sys[#i_Sys].Cnv_Level;

               IF "Settings_DB".ECnv_Sys[#i_Sys].Cnv_Level >= "Settings_DB".VTD_Sys[#i_Sys].Lowest_Level AND
                   "Settings_DB".ECnv_Sys[#i_Sys].Cnv_Level <= "Settings_DB".VTD_Sys[#i_Sys].Highest_Level AND //Leveled
                   "Control_DB".ECnv_Sys[#i_Sys].Cnv_Occupied AND //Econveyor occupied
                   NOT "Control_DB".ECnv_Sys[#i_Sys].Error AND //not error
                   NOT "Control_DB".ECnv_Sys[#i_Sys].Running AND //not error
                   ("Control_DB".LCnv_Sys[#i_Sys].Cnv_Level[#Level].Cnv1.Instruction.Inbound_Ready OR
                   "Control_DB".LCnv_Sys[#i_Sys].Cnv_Level[#Level].Cnv2.Instruction.Inbound_Ready) AND //conveyor not occupied
                   ("Control_DB".LCnv_Sys[#i_Sys].Cnv_Level[#Level].Cnv1.Mode = 2 OR
                   "Control_DB".LCnv_Sys[#i_Sys].Cnv_Level[#Level].Cnv1.Mode = 3 OR "Control_DB".LCnv_Sys[#i_Sys].Cnv_Level[#Level].Cnv2.Mode = 2 OR
                   "Control_DB".LCnv_Sys[#i_Sys].Cnv_Level[#Level].Cnv2.Mode = 3) AND //cnv1 or cnv 2 semi or auto mode
                   ("Control_DB".ECnv_Sys[#i_Sys].Mode = 2 OR "Control_DB".ECnv_Sys[#i_Sys].Mode = 3) THEN //Econveyor semi or auto mode 
                   "Control_DB".ECnv_Sys[#i_Sys].Instruction.Outbound_Ready := TRUE;
               ELSIF  NOT "Control_DB".ECnv_Sys[#i_Sys].Cnv_Occupied THEN  // // // // // // // // // // // // //last change
                   "Control_DB".ECnv_Sys[#i_Sys].Instruction.Outbound_Ready := FALSE;  // // // // // // // // // // // // //last change
               END_IF;


               //BUFFER CONVEYORS
               FOR #i_Lev := "Settings_DB".VTD_Sys[#i_Sys].Lowest_Level TO "Settings_DB".VTD_Sys[#i_Sys].Highest_Level DO
                   //CNV 1
                   IF "Control_DB".ECnv_Sys[#i_Sys].Instruction.Inbound_Ready AND
                       "Control_DB".VTD_Sys[#i_Sys].Current_Level = #i_Lev AND
                       (NOT "Control_DB".LCnv_Sys[#i_Sys].Cnv_Level[#i_Lev].Cnv2.Instruction.Transfer_in_Progress OR "Control_DB".VTD_Sys[#i_Sys].Current_Level = 1) AND
                       "Control_DB".LCnv_Sys[#i_Sys].Cnv_Level[#i_Lev].Cnv1.Cnv_Occupied AND
                       NOT "Control_DB".LCnv_Sys[#i_Sys].Cnv_Level[#i_Lev].Cnv1.Error AND NOT "Control_DB".LCnv_Sys[#i_Sys].Cnv_Level[#i_Lev].Cnv1.Running AND
                       ("Control_DB".LCnv_Sys[#i_Sys].Cnv_Level[#i_Lev].Cnv1.Mode = 2 OR "Control_DB".LCnv_Sys[#i_Sys].Cnv_Level[#i_Lev].Cnv1.Mode = 3) THEN
                       "Control_DB".LCnv_Sys[#i_Sys].Cnv_Level[#i_Lev].Cnv1.Instruction.Outbound_Ready := TRUE;
                   ELSIF  NOT "Control_DB".LCnv_Sys[#i_Sys].Cnv_Level[#i_Lev].Cnv1.Cnv_Occupied THEN  // // // // // // // // // // // // //last change
                       "Control_DB".LCnv_Sys[#i_Sys].Cnv_Level[#i_Lev].Cnv1.Instruction.Outbound_Ready := FALSE;  // // // // // // // // // // // // //last change
                   END_IF;

                   //CNV 2
                   IF ("Control_DB".ECnv_Sys[#i_Sys].Instruction.Inbound_Ready OR "Settings_DB".LCnv_Sys[#i_Sys].Cnv_Level[#i_Lev].Cnv2.Cnv_Level = 1) AND
                       ("Control_DB".VTD_Sys[#i_Sys].Current_Level = #i_Lev OR "Settings_DB".LCnv_Sys[#i_Sys].Cnv_Level[#i_Lev].Cnv2.Cnv_Level = 1) AND
                       (NOT "Control_DB".LCnv_Sys[#i_Sys].Cnv_Level[#i_Lev].Cnv1.Instruction.Transfer_in_Progress OR "Settings_DB".LCnv_Sys[#i_Sys].Cnv_Level[#i_Lev].Cnv2.Cnv_Level = 1) AND
                       "Control_DB".LCnv_Sys[#i_Sys].Cnv_Level[#i_Lev].Cnv2.Cnv_Occupied AND
                       NOT "Control_DB".LCnv_Sys[#i_Sys].Cnv_Level[#i_Lev].Cnv2.Error AND NOT "Control_DB".LCnv_Sys[#i_Sys].Cnv_Level[#i_Lev].Cnv2.Running AND
                       ("Control_DB".LCnv_Sys[#i_Sys].Cnv_Level[#i_Lev].Cnv2.Mode = 2 OR "Control_DB".LCnv_Sys[#i_Sys].Cnv_Level[#i_Lev].Cnv2.Mode = 3) THEN
                       "Control_DB".LCnv_Sys[#i_Sys].Cnv_Level[#i_Lev].Cnv2.Instruction.Outbound_Ready := TRUE;
                   ELSIF  NOT "Control_DB".LCnv_Sys[#i_Sys].Cnv_Level[#i_Lev].Cnv2.Cnv_Occupied THEN  // // // // // // // // // // // // //last change
                       "Control_DB".LCnv_Sys[#i_Sys].Cnv_Level[#i_Lev].Cnv2.Instruction.Outbound_Ready := FALSE;  // // // // // // // // // // // // //last change
                   END_IF;
               END_FOR;
           END_REGION

           REGION TRANSFER IN PROGRESS FOR EXTRACTOR CONVEYOR
               FOR #i_Lev := "Settings_DB".VTD_Sys[#i_Sys].Lowest_Level TO "Settings_DB".VTD_Sys[#i_Sys].Highest_Level DO
                   "Control_DB".ECnv_Sys[#i_Sys].Instruction.Transfer_in_Progress :=
                   ("Settings_DB".ECnv_Sys[#i_Sys].Cnv_Level = #i_Lev AND
                   "Control_DB".LCnv_Sys[#i_Sys].Cnv_Level[#i_Lev].Cnv1.Instruction.Transfer_in_Progress OR "Control_DB".LCnv_Sys[#i_Sys].Cnv_Level[#i_Lev].Cnv2.Instruction.Transfer_in_Progress);
               END_FOR;
           END_REGION
       END_FOR;

       IF "FirstScan" THEN
           "Time_1_Start_Buffers" := T#500MS;
           "Time_1_end_Buffers" := T#1S;
           "Time_2_Start_Buffers" := T#1S;
           "Time_2_End_Buffers" := T#1S_500MS;
           "Time_3_Buffers" := T#1S_500MS;

           "Time_1_Start_Ecnv" := T#1S700MS;
           "Time_1_end_Ecnv" := T#2S100MS;
           "Time_2_Start_Ecnv" := T#2S100MS;
           "Time_2_End_Ecnv" := T#2S_600MS;
           "Time_3_Ecnv" := T#2S_600MS;
       END_IF;
END_FUNCTION

FUNCTION "Bypass_FC" : Void   // FC62, SCL
{ S7_Optimized_Access := 'TRUE' }
VERSION : 0.1
// stored: AutoNumber true, IsIECCheckEnabled false, SetENOAutomatically false, UDAEnableTagReadback false
   VAR CONSTANT
      AUTO_RUNNING : UInt := 0;
      RTE_REQUESTED : UInt := 1;
      SAFE_BYPASS : UInt := 2;
      SAFE_TO_UNLOCK : UInt := 3;
      ACCESS_MANUAL_MODE : UInt := 4;
      READY_TO_RESET : UInt := 5;
      RESETTING : UInt := 6;
      READY_TO_RESTART : UInt := 7;
   END_VAR
BEGIN
   REGION LIGHT GUARD "Bypass"
       IF "FirstScan" THEN
           "MR_Delay_I" := T#1500mS;
           "MR_Delay_O" := T#1500mS;
       END_IF;

       // SYSTEM 1
       (*IF "Control_DB".LCnv_Sys[1].Cnv_Level[1].Cnv1.Running THEN //Running
           "Bypass".Remote_Panel_1."Light Guards CX101 - CH1" := TRUE; //Bypass light guard
           "Light_Guard_Bypass(1)" := FALSE; // Cancel HMI Command
       ELS*)IF "Control_DB".LCnv_Sys[1].Cnv_Level[1].Cnv1.Error AND "Light_Guard_Bypass(1)" THEN //Error and HMI command ON
           "Bypass".Remote_Panel_1."Light Guards CX101 - CH1" := TRUE; //Bypass light guard
       ELSIF NOT "Control_DB".LCnv_Sys[1].Cnv_Level[1].Cnv1.Running AND NOT "Control_DB".LCnv_Sys[1].Cnv_Level[1].Cnv1.Error AND "LIGHT GUARDS C1101 - CH1" THEN //Not Running and No error
           "Bypass".Remote_Panel_1."Light Guards CX101 - CH1" := FALSE; //Cancel bypass
       END_IF;

       (*IF "Control_DB".LCnv_Sys[1].Cnv_Level[1].Cnv2.Running THEN
           "Bypass".Remote_Panel_1."Light Guards CX201 - CH1" := TRUE;
           "Light_Guard_Bypass(1)" := FALSE;
       ELS*)IF "Control_DB".LCnv_Sys[1].Cnv_Level[1].Cnv2.Error AND "Light_Guard_Bypass(1)" THEN
           "Bypass".Remote_Panel_1."Light Guards CX201 - CH1" := TRUE;
       ELSIF NOT "Control_DB".LCnv_Sys[1].Cnv_Level[1].Cnv2.Running AND NOT "Control_DB".LCnv_Sys[1].Cnv_Level[1].Cnv2.Error AND "LIGHT GUARDS C1201 - CH1"THEN
           "Bypass".Remote_Panel_1."Light Guards CX201 - CH1" := FALSE;
       END_IF;

       //Request mute
       //Recognize starting pallet
       "R_Starting_Pallet_1"(CLK:= "DB_Receive_Data_From_Logistex".CNV_STATUS[1].%X6);
       IF "R_Starting_Pallet_1".Q AND "DB_Receive_Data_From_Logistex".J1310_Conv_Infeed.LGXTransferingInProgress THEN
           // Statement section IF
           "Starting_Pallet_1" := TRUE;

       ELSIF NOT "DB_Receive_Data_From_Logistex".J1310_Conv_Infeed.LGXTransferingInProgress OR "Control_DB".LCnv_Sys[1].Cnv_Level[1].Cnv1.Error THEN
           "Starting_Pallet_1" := FALSE;
       END_IF; 



       //Delay to start MR
       "T_MR_I_1".TON(IN := "DB_Receive_Data_From_Logistex".J1310_Conv_Infeed.LGXTransferingInProgress AND "Starting_Pallet_1",
                      PT := "MR_Delay_I",
                      Q => "MR_I_1");

       //INBOUND MATERIAL SELECTION
       IF "DB_Receive_Data_From_Logistex".J1310_Conv_Infeed.Pallet_ID[23] = 'U' THEN
           "Material_Selection_I_1" := FALSE;
       ELSIF "DB_Receive_Data_From_Logistex".J1310_Conv_Infeed.Pallet_ID[23] = 'E' THEN
           "Material_Selection_I_1" := TRUE;
       END_IF;

       //Delay to start MR
       "T_MR_O_1".TON(IN := "Control_DB".LCnv_Sys[1].Cnv_Level[1].Cnv2.SM_State = 40,
                      PT := "MR_Delay_O",
                      Q => "MR_O_1");

       //OUTBOUND MATERIAL SELECTION
       IF NOT "Control_DB".LCnv_Sys[1].Cnv_Level[1].Cnv2.Running AND "Control_DB".LCnv_Sys[1].Cnv_Level[1].Cnv2.Pallet_Type = 1 THEN
           "Material_Selection_O_1" := FALSE;
       ELSIF NOT "Control_DB".LCnv_Sys[1].Cnv_Level[1].Cnv2.Running AND "Control_DB".LCnv_Sys[1].Cnv_Level[1].Cnv2.Pallet_Type = 3 THEN
           "Material_Selection_O_1" := TRUE;
       END_IF;

       //SYSTEM 2
       (*IF "Control_DB".LCnv_Sys[2].Cnv_Level[1].Cnv1.Running THEN
           "Bypass".Remote_Panel_2."Light Guards CX101 - CH1" := TRUE;
           "Light_Guard_Bypass(2)" := FALSE;
       ELS*)IF "Control_DB".LCnv_Sys[2].Cnv_Level[1].Cnv1.Error AND "Light_Guard_Bypass(2)" THEN
           "Bypass".Remote_Panel_2."Light Guards CX101 - CH1" := TRUE;
       ELSIF NOT "Control_DB".LCnv_Sys[2].Cnv_Level[1].Cnv1.Running AND NOT "Control_DB".LCnv_Sys[2].Cnv_Level[1].Cnv1.Error AND "LIGHT GUARDS C2101 - CH1" THEN
           "Bypass".Remote_Panel_2."Light Guards CX101 - CH1" := FALSE;
       END_IF;

       (*IF "Control_DB".LCnv_Sys[2].Cnv_Level[1].Cnv2.Running THEN
           "Bypass".Remote_Panel_2."Light Guards CX201 - CH1" := TRUE;
           "Light_Guard_Bypass(2)" := FALSE;
       ELS*)IF "Control_DB".LCnv_Sys[2].Cnv_Level[1].Cnv2.Error AND "Light_Guard_Bypass(2)" THEN
           "Bypass".Remote_Panel_2."Light Guards CX201 - CH1" := TRUE;
       ELSIF NOT "Control_DB".LCnv_Sys[2].Cnv_Level[1].Cnv2.Running AND NOT "Control_DB".LCnv_Sys[2].Cnv_Level[1].Cnv2.Error AND "LIGHT GUARDS C2201 - CH1" THEN
           "Bypass".Remote_Panel_2."Light Guards CX201 - CH1" := FALSE;
       END_IF;

       //Request mute
       //Recognize starting pallet
       "R_Starting_Pallet_2"(CLK := "DB_Receive_Data_From_Logistex".CNV_STATUS[2].%X6);
       IF "R_Starting_Pallet_2".Q AND "DB_Receive_Data_From_Logistex".J1320_Conv_Infeed.LGXTransferingInProgress THEN
           // Statement section IF
           "Starting_Pallet_2" := TRUE;

       ELSIF NOT "DB_Receive_Data_From_Logistex".J1320_Conv_Infeed.LGXTransferingInProgress OR "Control_DB".LCnv_Sys[2].Cnv_Level[1].Cnv1.Error THEN
           "Starting_Pallet_2" := FALSE;
       END_IF;

       //Delay to start MR
       "T_MR_I_2".TON(IN := "DB_Receive_Data_From_Logistex".J1320_Conv_Infeed.LGXTransferingInProgress AND "Starting_Pallet_2",
                      PT := "MR_Delay_I",
                      Q => "MR_I_2");

       //INBOUND MATERIAL SELECTION
       IF "DB_Receive_Data_From_Logistex".J1320_Conv_Infeed.Pallet_ID[23] = 'U' THEN
           "Material_Selection_I_2" := FALSE;
       ELSIF "DB_Receive_Data_From_Logistex".J1320_Conv_Infeed.Pallet_ID[23] = 'E' THEN
           "Material_Selection_I_2" := TRUE;
       END_IF;

       //Delay to start MR
       "T_MR_O_2".TON(IN := "Control_DB".LCnv_Sys[2].Cnv_Level[1].Cnv2.SM_State = 40,
                      PT := "MR_Delay_O",
                      Q => "MR_O_2");

       //OUTBOUND MATERIAL SELECTION
       IF NOT "Control_DB".LCnv_Sys[2].Cnv_Level[1].Cnv2.Running AND "Control_DB".LCnv_Sys[2].Cnv_Level[1].Cnv2.Pallet_Type = 1 THEN
           "Material_Selection_O_2" := FALSE;
       ELSIF NOT "Control_DB".LCnv_Sys[2].Cnv_Level[1].Cnv2.Running AND "Control_DB".LCnv_Sys[2].Cnv_Level[1].Cnv2.Pallet_Type = 3 THEN
           "Material_Selection_O_2" := TRUE;
       END_IF;

       //SYSTEM 3
       (*IF "Control_DB".LCnv_Sys[3].Cnv_Level[1].Cnv1.Running THEN
           "Bypass".Remote_Panel_3."Light Guards CX101 - CH1" := TRUE;
           "Light_Guard_Bypass(3)" := FALSE;
       ELS*)IF "Control_DB".LCnv_Sys[3].Cnv_Level[1].Cnv1.Error AND "Light_Guard_Bypass(3)" THEN
           "Bypass".Remote_Panel_3."Light Guards CX101 - CH1" := TRUE;
       ELSIF NOT "Control_DB".LCnv_Sys[3].Cnv_Level[1].Cnv1.Running AND NOT "Control_DB".LCnv_Sys[3].Cnv_Level[1].Cnv1.Error AND "LIGHT GUARDS C3101 - CH1" THEN
           "Bypass".Remote_Panel_3."Light Guards CX101 - CH1" := FALSE;
       END_IF;

       (*IF "Control_DB".LCnv_Sys[3].Cnv_Level[1].Cnv2.Running THEN
           "Bypass".Remote_Panel_3."Light Guards CX201 - CH1" := TRUE;
           "Light_Guard_Bypass(3)" := FALSE;
       ELS*)IF "Control_DB".LCnv_Sys[3].Cnv_Level[1].Cnv2.Error AND "Light_Guard_Bypass(3)" THEN
           "Bypass".Remote_Panel_3."Light Guards CX201 - CH1" := TRUE;
       ELSIF NOT "Control_DB".LCnv_Sys[3].Cnv_Level[1].Cnv2.Running AND NOT "Control_DB".LCnv_Sys[3].Cnv_Level[1].Cnv2.Error AND "LIGHT GUARDS C3201 - CH1" THEN
           "Bypass".Remote_Panel_3."Light Guards CX201 - CH1" := FALSE;
       END_IF;

       //Request mute
       //Recognize starting pallet
       "R_Starting_Pallet_3"(CLK := "DB_Receive_Data_From_Logistex".CNV_STATUS[3].%X6);
       IF "R_Starting_Pallet_3".Q AND "DB_Receive_Data_From_Logistex".J1330_Conv_Infeed.LGXTransferingInProgress THEN
           // Statement section IF
           "Starting_Pallet_3" := TRUE;

       ELSIF NOT "DB_Receive_Data_From_Logistex".J1330_Conv_Infeed.LGXTransferingInProgress OR "Control_DB".LCnv_Sys[3].Cnv_Level[1].Cnv1.Error THEN
           "Starting_Pallet_3" := FALSE;
       END_IF;

       //Delay to start MR
       "T_MR_I_3".TON(IN := "DB_Receive_Data_From_Logistex".J1330_Conv_Infeed.LGXTransferingInProgress AND "Starting_Pallet_3",
                      PT := "MR_Delay_I",
                      Q => "MR_I_3");

       //INBOUND MATERIAL SELECTION
       IF "DB_Receive_Data_From_Logistex".J1330_Conv_Infeed.Pallet_ID[23] = 'U' THEN
           "Material_Selection_I_3" := FALSE;
       ELSIF "DB_Receive_Data_From_Logistex".J1330_Conv_Infeed.Pallet_ID[23] = 'E' THEN
           "Material_Selection_I_3" := TRUE;
       END_IF;

       //Delay to start MR
       "T_MR_O_3".TON(IN := "Control_DB".LCnv_Sys[3].Cnv_Level[1].Cnv2.SM_State = 40,
                      PT := "MR_Delay_O",
                      Q => "MR_O_3");

       //OUTBOUND MATERIAL SELECTION
       IF NOT "Control_DB".LCnv_Sys[3].Cnv_Level[1].Cnv2.Running AND "Control_DB".LCnv_Sys[3].Cnv_Level[1].Cnv2.Pallet_Type = 1 THEN
           "Material_Selection_O_3" := FALSE;
       ELSIF NOT "Control_DB".LCnv_Sys[3].Cnv_Level[1].Cnv2.Running AND "Control_DB".LCnv_Sys[3].Cnv_Level[1].Cnv2.Pallet_Type = 3 THEN
           "Material_Selection_O_3" := TRUE;
       END_IF;
   END_REGION ;

   REGION LIMIT SWITCHES
       REGION SYSTEM 1
           IF "VTD_System_Selected_HMI" = 1 THEN
               //OVERTRAVEL UP
               IF NOT "OVERTRAVEL UPPER LIMIT - CH1(1)" THEN
                   "Bypass".Remote_Panel_1.Overtravel_Upper_limit := "VTD_Upper_Overtravel_Bypass_HMI";
                   "T_Bypass_OUL_1".TON(IN := FALSE,
                                        PT := T#0S);
               ELSE
                   "T_Bypass_OUL_1".TON(IN := TRUE,
                                        PT := T#3S);
                   IF "T_Bypass_OUL_1".Q THEN
                       "Bypass".Remote_Panel_1.Overtravel_Upper_limit := "VTD_Upper_Overtravel_Bypass_HMI" := FALSE;
                   END_IF;
               END_IF;

               //LIMIT UP
               IF "VTD1 UPPER LIMIT" THEN
                   "Bypass".Remote_Panel_1.Upper_limit := "VTD_Upper_Limet_Bypass_HMI";
                   "T_Bypass_UL_1".TON(IN:=FALSE,
                                       PT:=T#0S);
               ELSE
                   "T_Bypass_UL_1".TON(IN := TRUE,
                                       PT := T#3S);
                   IF "T_Bypass_UL_1".Q THEN
                       "Bypass".Remote_Panel_1.Upper_limit := "VTD_Upper_Limet_Bypass_HMI" := FALSE;
                   END_IF;
               END_IF;

               //LIMIT DOWN
               IF "VTD1 LOWER LIMIT" THEN
                   "Bypass".Remote_Panel_1.Lower_limit := "VTD_Lower_Limit_Bypass_HMI";
                   "T_Bypass_LL_1".TON(IN:=FALSE,
                                       PT:=T#0S);
               ELSE
                   "T_Bypass_LL_1".TON(IN := TRUE,
                                       PT := T#3S);
                   IF "T_Bypass_LL_1".Q THEN
                       "Bypass".Remote_Panel_1.Lower_limit := "VTD_Lower_Limit_Bypass_HMI" := FALSE;
                   END_IF;
               END_IF;

               //OVERTRAVEL DOWN
               IF NOT "OVERTRAVEL LOWER LIMIT - CH1(1)" THEN
                   "Bypass".Remote_Panel_1.Overtravel_Lower_limit := "VTD_Lower_Overtravel_Bypass_HMI";
                   "T_Bypass_OLL_1".TON(IN:=FALSE,
                                        PT:=T#0S);
               ELSE
                   "T_Bypass_OLL_1".TON(IN := TRUE,
                                        PT := T#3S);
                   IF "T_Bypass_OLL_1".Q THEN
                       "Bypass".Remote_Panel_1.Overtravel_Lower_limit := "VTD_Lower_Overtravel_Bypass_HMI" := FALSE;
                   END_IF;
               END_IF;

               //CHAIN SLACK 1
               IF "Chain Slack 1 - CH1(1)" THEN
                   "Bypass".Remote_Panel_1.Chain_Slack_1 := "Chain_Slack_1_Bypass_HMI";
               ELSE
                   "Bypass".Remote_Panel_1.Chain_Slack_1 := "Chain_Slack_1_Bypass_HMI" := FALSE;
               END_IF;

               //CHAIN SLACK 2
               IF "Chain Slack 2 - CH1(1)" THEN
                   "Bypass".Remote_Panel_1.Chain_Slack_2 := "Chain_Slack_2_Bypass_HMI";
               ELSE
                   "Bypass".Remote_Panel_1.Chain_Slack_2 := "Chain_Slack_2_Bypass_HMI" := FALSE;
               END_IF;

               //CHAIN SLACK 3
               IF "Chain Slack 3 - CH1(1)" THEN
                   "Bypass".Remote_Panel_1.Chain_Slack_3 := "Chain_Slack_3_Bypass_HMI";
               ELSE
                   "Bypass".Remote_Panel_1.Chain_Slack_3 := "Chain_Slack_3_Bypass_HMI" := FALSE;
               END_IF;

               //CHAIN SLACK 4
               IF "Chain Slack 4 - CH1(1)" THEN
                   "Bypass".Remote_Panel_1.Chain_Slack_4 := "Chain_Slack_4_Bypass_HMI";
               ELSE
                   "Bypass".Remote_Panel_1.Chain_Slack_4 := "Chain_Slack_4_Bypass_HMI" := FALSE;
               END_IF;
           END_IF;
       END_REGION ;

       REGION SYSTEM 2
           IF "VTD_System_Selected_HMI" = 2 THEN
               //OVERTRAVEL UP
               IF NOT "OVERTRAVEL UPPER LIMIT - CH1(2)" THEN
                   "Bypass".Remote_Panel_2.Overtravel_Upper_limit := "VTD_Upper_Overtravel_Bypass_HMI";
                   "T_Bypass_OUL_2".TON(IN := FALSE,
                                        PT := T#0S);
               ELSE
                   "T_Bypass_OUL_2".TON(IN := TRUE,
                                        PT := T#3S);
                   IF "T_Bypass_OUL_2".Q THEN
                       "Bypass".Remote_Panel_2.Overtravel_Upper_limit := "VTD_Upper_Overtravel_Bypass_HMI" := FALSE;
                   END_IF;
               END_IF;

               //LIMIT UP
               IF "VTD2 UPPER LIMIT" THEN
                   "Bypass".Remote_Panel_2.Upper_limit := "VTD_Upper_Limet_Bypass_HMI";
                   "T_Bypass_UL_2".TON(IN := FALSE,
                                       PT := T#0S);
               ELSE
                   "T_Bypass_UL_2".TON(IN := TRUE,
                                       PT := T#3S);
                   IF "T_Bypass_UL_2".Q THEN
                       "Bypass".Remote_Panel_2.Upper_limit := "VTD_Upper_Limet_Bypass_HMI" := FALSE;
                   END_IF;
               END_IF;

               //LIMIT DOWN
               IF "VTD2 LOWER LIMIT" THEN
                   "Bypass".Remote_Panel_2.Lower_limit := "VTD_Lower_Limit_Bypass_HMI";
                   "T_Bypass_LL_2".TON(IN := FALSE,
                                       PT := T#0S);
               ELSE
                   "T_Bypass_LL_2".TON(IN := TRUE,
                                       PT := T#3S);
                   IF "T_Bypass_LL_2".Q THEN
                       "Bypass".Remote_Panel_2.Lower_limit := "VTD_Lower_Limit_Bypass_HMI" := FALSE;
                   END_IF;
               END_IF;

               //OVERTRAVEL DOWN
               IF NOT "OVERTRAVEL LOWER LIMIT - CH1(2)" THEN
                   "Bypass".Remote_Panel_2.Overtravel_Lower_limit := "VTD_Lower_Overtravel_Bypass_HMI";
                   "T_Bypass_OLL_2".TON(IN := FALSE,
                                        PT := T#0S);
               ELSE
                   "T_Bypass_OLL_2".TON(IN := TRUE,
                                        PT := T#3S);
                   IF "T_Bypass_OLL_2".Q THEN
                       "Bypass".Remote_Panel_2.Overtravel_Lower_limit := "VTD_Lower_Overtravel_Bypass_HMI" := FALSE;
                   END_IF;
               END_IF;

               //CHAIN SLACK 1
               IF "Chain Slack 1 - CH1(2)" THEN
                   "Bypass".Remote_Panel_2.Chain_Slack_1 := "Chain_Slack_1_Bypass_HMI";
               ELSE
                   "Bypass".Remote_Panel_2.Chain_Slack_1 := "Chain_Slack_1_Bypass_HMI" := FALSE;
               END_IF;

               //CHAIN SLACK 2
               IF "Chain Slack 2 - CH1(2)" THEN
                   "Bypass".Remote_Panel_2.Chain_Slack_2 := "Chain_Slack_2_Bypass_HMI";
               ELSE
                   "Bypass".Remote_Panel_2.Chain_Slack_2 := "Chain_Slack_2_Bypass_HMI" := FALSE;
               END_IF;

               //CHAIN SLACK 3
               IF "Chain Slack 3 - CH1(2)" THEN
                   "Bypass".Remote_Panel_2.Chain_Slack_3 := "Chain_Slack_3_Bypass_HMI";
               ELSE
                   "Bypass".Remote_Panel_2.Chain_Slack_3 := "Chain_Slack_3_Bypass_HMI" := FALSE;
               END_IF;

               //CHAIN SLACK 4
               IF "Chain Slack 4 - CH1(2)" THEN
                   "Bypass".Remote_Panel_2.Chain_Slack_4 := "Chain_Slack_4_Bypass_HMI";
               ELSE
                   "Bypass".Remote_Panel_2.Chain_Slack_4 := "Chain_Slack_4_Bypass_HMI" := FALSE;
               END_IF;
           END_IF;
       END_REGION ;

       REGION SYSTEM 3
           IF "VTD_System_Selected_HMI" = 3 THEN
               //OVERTRAVEL UP
               IF NOT "OVERTRAVEL UPPER LIMIT - CH1(3)" THEN
                   "Bypass".Remote_Panel_3.Overtravel_Upper_limit := "VTD_Upper_Overtravel_Bypass_HMI";
                   "T_Bypass_OUL_3".TON(IN := FALSE,
                                        PT := T#0S);
               ELSE
                   "T_Bypass_OUL_3".TON(IN := TRUE,
                                        PT := T#3S);
                   IF "T_Bypass_OUL_3".Q THEN
                       "Bypass".Remote_Panel_3.Overtravel_Upper_limit := "VTD_Upper_Overtravel_Bypass_HMI" := FALSE;
                   END_IF;
               END_IF;

               //LIMIT UP
               IF "VTD3 UPPER LIMIT" THEN
                   "Bypass".Remote_Panel_3.Upper_limit := "VTD_Upper_Limet_Bypass_HMI";
                   "T_Bypass_UL_3".TON(IN := FALSE,
                                       PT := T#0S);
               ELSE
                   "T_Bypass_UL_3".TON(IN := TRUE,
                                       PT := T#3S);
                   IF "T_Bypass_UL_3".Q THEN
                       "Bypass".Remote_Panel_3.Upper_limit := "VTD_Upper_Limet_Bypass_HMI" := FALSE;
                   END_IF;
               END_IF;

               //LIMIT DOWN
               IF "VTD3 LOWER LIMIT" THEN
                   "Bypass".Remote_Panel_3.Lower_limit := "VTD_Lower_Limit_Bypass_HMI";
                   "T_Bypass_LL_3".TON(IN := FALSE,
                                       PT := T#0S);
               ELSE
                   "T_Bypass_LL_3".TON(IN := TRUE,
                                       PT := T#3S);
                   IF "T_Bypass_LL_3".Q THEN
                       "Bypass".Remote_Panel_3.Lower_limit := "VTD_Lower_Limit_Bypass_HMI" := FALSE;
                   END_IF;
               END_IF;

               //OVERTRAVEL DOWN
               IF NOT "OVERTRAVEL LOWER LIMIT - CH1(3)" THEN
                   "Bypass".Remote_Panel_3.Overtravel_Lower_limit := "VTD_Lower_Overtravel_Bypass_HMI";
                   "T_Bypass_OLL_3".TON(IN := FALSE,
                                        PT := T#0S);
               ELSE
                   "T_Bypass_OLL_3".TON(IN := TRUE,
                                        PT := T#3S);
                   IF "T_Bypass_OLL_3".Q THEN
                       "Bypass".Remote_Panel_3.Overtravel_Lower_limit := "VTD_Lower_Overtravel_Bypass_HMI" := FALSE;
                   END_IF;
               END_IF;

               //CHAIN SLACK 1
               IF "Chain Slack 1 - CH1(3)" THEN
                   "Bypass".Remote_Panel_3.Chain_Slack_1 := "Chain_Slack_1_Bypass_HMI";
               ELSE
                   "Bypass".Remote_Panel_3.Chain_Slack_1 := "Chain_Slack_1_Bypass_HMI" := FALSE;
               END_IF;

               //CHAIN SLACK 2
               IF "Chain Slack 2 - CH1(3)" THEN
                   "Bypass".Remote_Panel_3.Chain_Slack_2 := "Chain_Slack_2_Bypass_HMI";
               ELSE
                   "Bypass".Remote_Panel_3.Chain_Slack_2 := "Chain_Slack_2_Bypass_HMI" := FALSE;
               END_IF;

               //CHAIN SLACK 3
               IF "Chain Slack 3 - CH1(3)" THEN
                   "Bypass".Remote_Panel_3.Chain_Slack_3 := "Chain_Slack_3_Bypass_HMI";
               ELSE
                   "Bypass".Remote_Panel_3.Chain_Slack_3 := "Chain_Slack_3_Bypass_HMI" := FALSE;
               END_IF;

               //CHAIN SLACK 4
               IF "Chain Slack 4 - CH1(3)" THEN
                   "Bypass".Remote_Panel_3.Chain_Slack_4 := "Chain_Slack_4_Bypass_HMI";
               ELSE
                   "Bypass".Remote_Panel_3.Chain_Slack_4 := "Chain_Slack_4_Bypass_HMI" := FALSE;
               END_IF;
           END_IF;
       END_REGION ;

       REGION SYSTEM 4
           IF "VTD_System_Selected_HMI" = 4 THEN
               //OVERTRAVEL UP
               IF NOT "OVERTRAVEL UPPER LIMIT - CH1(4)" THEN
                   "Bypass".Remote_Panel_4.Overtravel_Upper_limit := "VTD_Upper_Overtravel_Bypass_HMI";
                   "T_Bypass_OUL_4".TON(IN := FALSE,
                                        PT := T#0S);
               ELSE
                   "T_Bypass_OUL_4".TON(IN := TRUE,
                                        PT := T#3S);
                   IF "T_Bypass_OUL_4".Q THEN
                       "Bypass".Remote_Panel_4.Overtravel_Upper_limit := "VTD_Upper_Overtravel_Bypass_HMI" := FALSE;
                   END_IF;
               END_IF;

               //LIMIT UP
               IF "VTD4 UPPER LIMIT" THEN
                   "Bypass".Remote_Panel_4.Upper_limit := "VTD_Upper_Limet_Bypass_HMI";
                   "T_Bypass_UL_4".TON(IN := FALSE,
                                       PT := T#0S);
               ELSE
                   "T_Bypass_UL_4".TON(IN := TRUE,
                                       PT := T#3S);
                   IF "T_Bypass_UL_4".Q THEN
                       "Bypass".Remote_Panel_4.Upper_limit := "VTD_Upper_Limet_Bypass_HMI" := FALSE;
                   END_IF;
               END_IF;

               //LIMIT DOWN
               IF "VTD4 LOWER LIMIT" THEN
                   "Bypass".Remote_Panel_4.Lower_limit := "VTD_Lower_Limit_Bypass_HMI";
                   "T_Bypass_LL_4".TON(IN := FALSE,
                                       PT := T#0S);
               ELSE
                   "T_Bypass_LL_4".TON(IN := TRUE,
                                       PT := T#3S);
                   IF "T_Bypass_LL_4".Q THEN
                       "Bypass".Remote_Panel_4.Lower_limit := "VTD_Lower_Limit_Bypass_HMI" := FALSE;
                   END_IF;
               END_IF;

               //OVERTRAVEL DOWN
               IF NOT "OVERTRAVEL LOWER LIMIT - CH1(4)" THEN
                   "Bypass".Remote_Panel_4.Overtravel_Lower_limit := "VTD_Lower_Overtravel_Bypass_HMI";
                   "T_Bypass_OLL_4".TON(IN := FALSE,
                                        PT := T#0S);
               ELSE
                   "T_Bypass_OLL_4".TON(IN := TRUE,
                                        PT := T#3S);
                   IF "T_Bypass_OLL_4".Q THEN
                       "Bypass".Remote_Panel_4.Overtravel_Lower_limit := "VTD_Lower_Overtravel_Bypass_HMI" := FALSE;
                   END_IF;
               END_IF;

               //CHAIN SLACK 1
               IF "Chain Slack 1 - CH1(4)" THEN
                   "Bypass".Remote_Panel_4.Chain_Slack_1 := "Chain_Slack_1_Bypass_HMI";
               ELSE
                   "Bypass".Remote_Panel_4.Chain_Slack_1 := "Chain_Slack_1_Bypass_HMI" := FALSE;
               END_IF;

               //CHAIN SLACK 2
               IF "Chain Slack 2 - CH1(4)" THEN
                   "Bypass".Remote_Panel_4.Chain_Slack_2 := "Chain_Slack_2_Bypass_HMI";
               ELSE
                   "Bypass".Remote_Panel_4.Chain_Slack_2 := "Chain_Slack_2_Bypass_HMI" := FALSE;
               END_IF;

               //CHAIN SLACK 3
               IF "Chain Slack 3 - CH1(4)" THEN
                   "Bypass".Remote_Panel_4.Chain_Slack_3 := "Chain_Slack_3_Bypass_HMI";
               ELSE
                   "Bypass".Remote_Panel_4.Chain_Slack_3 := "Chain_Slack_3_Bypass_HMI" := FALSE;
               END_IF;

               //CHAIN SLACK 4
               IF "Chain Slack 4 - CH1(4)" THEN
                   "Bypass".Remote_Panel_4.Chain_Slack_4 := "Chain_Slack_4_Bypass_HMI";
               ELSE
                   "Bypass".Remote_Panel_4.Chain_Slack_4 := "Chain_Slack_4_Bypass_HMI" := FALSE;
               END_IF;
           END_IF;
       END_REGION ;

       REGION SYSTEM 5
           IF "VTD_System_Selected_HMI" = 5 THEN
               //OVERTRAVEL UP
               IF NOT "OVERTRAVEL UPPER LIMIT - CH1(5)" THEN
                   "Bypass".Remote_Panel_5.Overtravel_Upper_limit := "VTD_Upper_Overtravel_Bypass_HMI";
                   "T_Bypass_OUL_5".TON(IN := FALSE,
                                        PT := T#0S);
               ELSE
                   "T_Bypass_OUL_5".TON(IN := TRUE,
                                        PT := T#3S);
                   IF "T_Bypass_OUL_5".Q THEN
                       "Bypass".Remote_Panel_5.Overtravel_Upper_limit := "VTD_Upper_Overtravel_Bypass_HMI" := FALSE;
                   END_IF;
               END_IF;

               //LIMIT UP
               IF "VTD5 UPPER LIMIT" THEN
                   "Bypass".Remote_Panel_5.Upper_limit := "VTD_Upper_Limet_Bypass_HMI";
                   "T_Bypass_UL_5".TON(IN := FALSE,
                                       PT := T#0S);
               ELSE
                   "T_Bypass_UL_5".TON(IN := TRUE,
                                       PT := T#3S);
                   IF "T_Bypass_UL_5".Q THEN
                       "Bypass".Remote_Panel_5.Upper_limit := "VTD_Upper_Limet_Bypass_HMI" := FALSE;
                   END_IF;
               END_IF;

               //LIMIT DOWN
               IF "VTD5 LOWER LIMIT" THEN
                   "Bypass".Remote_Panel_5.Lower_limit := "VTD_Lower_Limit_Bypass_HMI";
                   "T_Bypass_LL_5".TON(IN := FALSE,
                                       PT := T#0S);
               ELSE
                   "T_Bypass_LL_5".TON(IN := TRUE,
                                       PT := T#3S);
                   IF "T_Bypass_LL_5".Q THEN
                       "Bypass".Remote_Panel_5.Lower_limit := "VTD_Lower_Limit_Bypass_HMI" := FALSE;
                   END_IF;
               END_IF;

               //OVERTRAVEL DOWN
               IF NOT "OVERTRAVEL LOWER LIMIT - CH1(5)" THEN
                   "Bypass".Remote_Panel_5.Overtravel_Lower_limit := "VTD_Lower_Overtravel_Bypass_HMI";
                   "T_Bypass_OLL_5".TON(IN := FALSE,
                                        PT := T#0S);
               ELSE
                   "T_Bypass_OLL_5".TON(IN := TRUE,
                                        PT := T#3S);
                   IF "T_Bypass_OLL_5".Q THEN
                       "Bypass".Remote_Panel_5.Overtravel_Lower_limit := "VTD_Lower_Overtravel_Bypass_HMI" := FALSE;
                   END_IF;
               END_IF;

               //CHAIN SLACK 1
               IF "Chain Slack 1 - CH1(5)" THEN
                   "Bypass".Remote_Panel_5.Chain_Slack_1 := "Chain_Slack_1_Bypass_HMI";
               ELSE
                   "Bypass".Remote_Panel_5.Chain_Slack_1 := "Chain_Slack_1_Bypass_HMI" := FALSE;
               END_IF;

               //CHAIN SLACK 2
               IF "Chain Slack 2 - CH1(5)" THEN
                   "Bypass".Remote_Panel_5.Chain_Slack_2 := "Chain_Slack_2_Bypass_HMI";
               ELSE
                   "Bypass".Remote_Panel_5.Chain_Slack_2 := "Chain_Slack_2_Bypass_HMI" := FALSE;
               END_IF;

               //CHAIN SLACK 3
               IF "Chain Slack 3 - CH1(5)" THEN
                   "Bypass".Remote_Panel_5.Chain_Slack_3 := "Chain_Slack_3_Bypass_HMI";
               ELSE
                   "Bypass".Remote_Panel_5.Chain_Slack_3 := "Chain_Slack_3_Bypass_HMI" := FALSE;
               END_IF;

               //CHAIN SLACK 4
               IF "Chain Slack 4 - CH1(5)" THEN
                   "Bypass".Remote_Panel_5.Chain_Slack_4 := "Chain_Slack_4_Bypass_HMI";
               ELSE
                   "Bypass".Remote_Panel_5.Chain_Slack_4 := "Chain_Slack_4_Bypass_HMI" := FALSE;
               END_IF;
           END_IF;
       END_REGION ;
   END_REGION

   REGION SAFETY GATES
           //SYSTEM 1
           // GATE 1
           IF "GateAccess_Station_FB_DB_1".ModeManager.CurrentState > #RTE_REQUESTED AND
               "GateAccess_Station_FB_DB_1".ModeManager.CurrentState < #READY_TO_RESTART THEN
               "Bypass".Remote_Panel_1.Gate_1 := TRUE;
               "Bypass".Remote_Panel_1.Lock_Secured_1 := TRUE;
           // ELSE
           //     "Bypass".Remote_Panel_1.Gate_1 := FALSE;
           //     "Bypass".Remote_Panel_1.Lock_Secured_1 := FALSE;
           END_IF;

           //GATE 2
           IF "GateAccess_Station_FB_DB_2".ModeManager.CurrentState > #RTE_REQUESTED AND
               "GateAccess_Station_FB_DB_2".ModeManager.CurrentState < #READY_TO_RESTART THEN
               "Bypass".Remote_Panel_1.Gate_2 := TRUE;
               "Bypass".Remote_Panel_1.Lock_Secured_2 := TRUE;
           // ELSE
           //     "Bypass".Remote_Panel_1.Gate_2 := FALSE;
           //     "Bypass".Remote_Panel_1.Lock_Secured_2 := FALSE;
           END_IF;

           //SYSTEM 2
           //GATE 1
           IF "GateAccess_Station_FB_DB_3".ModeManager.CurrentState > #RTE_REQUESTED AND
               "GateAccess_Station_FB_DB_3".ModeManager.CurrentState < #READY_TO_RESTART THEN
               "Bypass".Remote_Panel_2.Gate_1 := TRUE;
               "Bypass".Remote_Panel_2.Lock_Secured_1 := TRUE;
           ELSE
               "Bypass".Remote_Panel_2.Gate_1 := FALSE;
               "Bypass".Remote_Panel_2.Lock_Secured_1 := FALSE;
           END_IF;

           //GATE 2
           IF "GateAccess_Station_FB_DB_4".ModeManager.CurrentState > #RTE_REQUESTED AND
               "GateAccess_Station_FB_DB_4".ModeManager.CurrentState < #READY_TO_RESTART THEN
               "Bypass".Remote_Panel_2.Gate_2 := TRUE;
               "Bypass".Remote_Panel_2.Lock_Secured_2 := TRUE;
           ELSE
               "Bypass".Remote_Panel_2.Gate_2 := FALSE;
               "Bypass".Remote_Panel_2.Lock_Secured_2 := FALSE;
           END_IF;

           //SYSTEM 3
           //GATE 1
           IF "GateAccess_Station_FB_DB_5".ModeManager.CurrentState > #RTE_REQUESTED AND
               "GateAccess_Station_FB_DB_5".ModeManager.CurrentState < #READY_TO_RESTART THEN
               "Bypass".Remote_Panel_3.Gate_1 := TRUE;
               "Bypass".Remote_Panel_3.Lock_Secured_1 := TRUE;
           ELSE
               "Bypass".Remote_Panel_3.Gate_1 := FALSE;
               "Bypass".Remote_Panel_3.Lock_Secured_1 := FALSE;
           END_IF;

           //GATE 2
           IF "GateAccess_Station_FB_DB_6".ModeManager.CurrentState > #RTE_REQUESTED AND
               "GateAccess_Station_FB_DB_6".ModeManager.CurrentState < #READY_TO_RESTART THEN
               "Bypass".Remote_Panel_3.Gate_2 := TRUE;
               "Bypass".Remote_Panel_3.Lock_Secured_2 := TRUE;
           ELSE
               "Bypass".Remote_Panel_3.Gate_2 := FALSE;
               "Bypass".Remote_Panel_3.Lock_Secured_2 := FALSE;
           END_IF;

           //SYSTEM 4
           //GATE 1
           IF "GateAccess_Station_FB_DB_9".ModeManager.CurrentState > #RTE_REQUESTED AND
               "GateAccess_Station_FB_DB_9".ModeManager.CurrentState < #READY_TO_RESTART THEN
               "Bypass".Remote_Panel_4.Gate_1 := TRUE;
               "Bypass".Remote_Panel_4.Lock_Secured_1 := TRUE;
           ELSE
               "Bypass".Remote_Panel_4.Gate_1 := FALSE;
               "Bypass".Remote_Panel_4.Lock_Secured_1 := FALSE;
           END_IF;

           //SYSTEM 5
           //GATE 1
           IF "GateAccess_Station_FB_DB_10".ModeManager.CurrentState > #RTE_REQUESTED AND
               "GateAccess_Station_FB_DB_10".ModeManager.CurrentState < #READY_TO_RESTART THEN
               "Bypass".Remote_Panel_5.Gate_1 := TRUE;
               "Bypass".Remote_Panel_5.Lock_Secured_1 := TRUE;
           ELSE
               "Bypass".Remote_Panel_5.Gate_1 := FALSE;
               "Bypass".Remote_Panel_5.Lock_Secured_1 := FALSE;
           END_IF;

           //Left side
           //LEVEL 1
           IF "GateAccess_Station_FB_DB_7".ModeManager.CurrentState > #RTE_REQUESTED AND
               "GateAccess_Station_FB_DB_7".ModeManager.CurrentState < #READY_TO_RESTART THEN
               "Bypass".Main_Panel.Lock_Secured_7 := TRUE;
           ELSE
               "Bypass".Main_Panel.Lock_Secured_7 := FALSE;
           END_IF;

           //LEVEL 2
           IF "GateAccess_Station_FB_DB_8".ModeManager.CurrentState > #RTE_REQUESTED AND
               "GateAccess_Station_FB_DB_8".ModeManager.CurrentState < #READY_TO_RESTART THEN
               "Bypass".Main_Panel.Lock_Secured_8 := TRUE;
           ELSE
               "Bypass".Main_Panel.Lock_Secured_8 := FALSE;
           END_IF;

           //Right side
           //LEVEL 1
           IF "GateAccess_Station_FB_DB_12".ModeManager.CurrentState > #RTE_REQUESTED AND
               "GateAccess_Station_FB_DB_12".ModeManager.CurrentState < #READY_TO_RESTART THEN
               "Bypass".Main_Panel.Lock_Secured_12 := TRUE;
           ELSE
               "Bypass".Main_Panel.Lock_Secured_12 := FALSE;
           END_IF;

           //LEVEL 2
           IF "GateAccess_Station_FB_DB_11".ModeManager.CurrentState > #RTE_REQUESTED AND
               "GateAccess_Station_FB_DB_11".ModeManager.CurrentState < #READY_TO_RESTART THEN
               "Bypass".Main_Panel.Lock_Secured_11 := TRUE;
           ELSE
               "Bypass".Main_Panel.Lock_Secured_11 := FALSE;
           END_IF;
   END_REGION;
END_FUNCTION

FUNCTION "Local_Mode_FC" : Bool   // FC67, SCL
{ S7_Optimized_Access := 'TRUE' }
VERSION : 0.1
// stored: AutoNumber true, IsIECCheckEnabled false, SetENOAutomatically false, UDAEnableTagReadback false
   VAR_INPUT
      HMI_Box_Connected : Int;
      Rem_Loc_Keys : Array[1..5] of "Level_Keys_UDT";
   END_VAR
   VAR_TEMP
      System : UInt;
      Level : UInt;
   END_VAR
BEGIN
   #System := #HMI_Box_Connected / 10;
   #Level := #HMI_Box_Connected MOD 10;
   IF #System <> 0 AND #Level <> 0 THEN
       #Local_Mode_FC := #Rem_Loc_Keys[#System].Level[#Level];
   ELSE
       #Local_Mode_FC := FALSE;
   END_IF;
END_FUNCTION

FUNCTION_BLOCK "VTD_FB"   // FB18, SCL
{ S7_Optimized_Access := 'TRUE' }
VERSION : 0.1
// stored: AutoNumber true, IsIECCheckEnabled false, IsRetainMemResEnabled false, MemoryReserve 100, SetENOAutomatically false, UDAEnableTagReadback false
   VAR_INPUT
      System_no : UInt;
      Safety_OK_Delayed : Bool;
      Safety_OK : Bool;
      Cnv_Sensors : "Cnv_Inputs";
      VTD_Settings : "VTD_Settings";
      Bypass_LP : Bool;
      Bypass : "Safety_Bypass_RemotePanel";
   END_VAR
   VAR_IN_OUT
      VTD_Control : "VTD_Control";
      SinaSpeed : SinaSpeed;
      LE_Bypass_HMI : Bool;
   END_VAR
   VAR
      State : UInt;
      Last_State : UInt;
      I_State : UInt;
      LD_Timer_1 : TON_TIME;
      LD_Timer : TON_TIME;
      DP_Timer { S7_SetPoint := 'True'} : TON_TIME;
      Watchdog { S7_SetPoint := 'True'} : TON_TIME;
      CS_TImer { S7_SetPoint := 'True'} : TON_TIME;
      Interlock_Timer { S7_SetPoint := 'True'} : TON_TIME;
      MainSetpoint : Int;
      Position_Offset : Real;
      ChangeToLow : Array[1..4] of DInt;
      DestPosition : Real;
      SetUpSpeed : UInt;
      LevelBelowExtractor : UInt := 1;
      IEC_Timer_0_Instance { S7_SetPoint := 'True'} : TON_TIME;
      DestinationLevel : UInt;
      CurrentlLevel : UInt;
      VTD_ID_Decoded { ExternalAccessible := 'False'; ExternalVisible := 'False'; ExternalWritable := 'False'} : "ID_Decoded";
      Cnv_ID_Decoded { ExternalAccessible := 'False'; ExternalVisible := 'False'; ExternalWritable := 'False'} : Array[1..2] of "ID_Decoded";
      IEC_Timer_0_Instance_1 { S7_SetPoint := 'True'} : TON_TIME;
      IEC_Timer_0_Instance_2 { S7_SetPoint := 'True'} : TON_TIME;
      VTD_ControlInstructionTask_ID_Old : Int;
      R_Execulte { S7_SetPoint := 'True'} : R_TRIG;
      R_AutomatcMode { S7_SetPoint := 'True'} : R_TRIG;
      T_Encoders_Difference { S7_SetPoint := 'True'} : TON_TIME;
      T_LE_Error { S7_SetPoint := 'True'} : TON_TIME;
      T_Setpoint_Delay { S7_SetPoint := 'True'} : TON_TIME;
      Distance_mm : Real;
      TravelTime_s : UInt;
      LE_Prev_mm : Real;
      DeltaPos_mm : Real;
      SampleTime_s : Real := 0.1;
      VTDSpeed_mm_s : Real;
      T_Speed { S7_SetPoint := 'True'} : TON_TIME;
      Speed_mm_per_percent : Real := 8.0;
      Speed_mm_s { ExternalAccessible := 'False'; ExternalVisible := 'False'; ExternalWritable := 'False'} : Real;
      TravelTime_ms { ExternalAccessible := 'False'; ExternalVisible := 'False'; ExternalWritable := 'False'} : UInt;
      Watchdog_PT { ExternalAccessible := 'False'; ExternalVisible := 'False'; ExternalWritable := 'False'} : Time;
      Stopper_Extend_Timer { S7_SetPoint := 'True'} : TON_TIME;
      T_LE_read_0 { S7_SetPoint := 'True'} : TON_TIME;
   END_VAR
   VAR_TEMP
      Level_Accuracy : String;
      i : UInt;
      Upper_limit : Bool;
      Ultimate_SlowDown : Bool;
      Ultimate_Creep : Bool;
      Lower_Limit : Bool;
      Level_Detect : Bool;
      Level_Detect1 : Bool;
      Level_Detect2 : Bool;
      DP2_Extended : Bool;
      DP2_Retracted : Bool;
      DP1_Extended : Bool;
      DP1_Retracted : Bool;
      Chain_Slack_1 : Bool;
      Chain_Slack_2 : Bool;
      Chain_Slack_3 : Bool;
      Chain_Slack_4 : Bool;
      Shuttle_Detect1 : Bool;
      Shuttle_Detect2 : Bool;
      DP1_Retract : Bool;
      DP1_Extend : Bool;
      DP2_Retract : Bool;
      DP2_Extend : Bool;
      Cnvs1_NotExtended : Bool;
      Cnvs2_NotExtended : Bool;
      Stoppers_NotExtended : Bool;
      MainSetpoint1 : Int;
      HMI_Reset : Bool;
      ConfigAxis : Word;
   END_VAR
   VAR CONSTANT
      EMPTY : USInt := 0;
      CHEP : USInt := 1;
      "EURO LEFT" : USInt := 2;
      "EURO RIGHT" : USInt := 3;
      "EURO CENTER" : USInt := 4;
      UNKNOWN : USInt := 5;
   END_VAR
BEGIN
   //Execute
   #R_Execulte(CLK := #VTD_Control.Instruction.Execulte);

   IF #VTD_Control.Mode = 3 THEN
       #VTD_Control.Instruction.Enable := TRUE;
   END_IF;

   #VTD_Control.Enabled := #VTD_Control.Instruction.Enable;

   #VTD_Control.Mode := #VTD_Control.Instruction.Mode_Change;

   IF NOT #VTD_Control.Enabled AND NOT #VTD_Control.Error THEN
       #State := 0;
   END_IF;

   //MANUAL MODE
   IF (#VTD_Control.Mode = 1 OR #VTD_Control.Mode = 5) AND NOT #VTD_Control.Error AND #VTD_Control.Enabled THEN
       #State := 500;
   END_IF;

   (*
   TODO:

   Mode select is done via the HMI. Might add external mode select switches.

           Mode select mask:
           0: Disabled
           1: Manual
           2: Semi-Auto
           3: Auto
           4: Teach
           5: Maintenance

   Device ID Format: XXYYZZ    
   XX = Device type   
       01   VTD
       10  Cnv_Front_of_VTD
       11  Cnv_Rear_of_VTD
       12  Cnv_On_Extractor
       20  Safety_Stop_Front_of_VTD
       21  Safety_Stop_Rear_of_VTD
   YY = Floor   
   ZZ = VTD Connected to 
   *)

   REGION Sensor allocations
       //Assign inputs to local vars
       #Upper_limit := #VTD_Control.Inputs.Upper_limit;
       #Ultimate_SlowDown := #VTD_Control.Inputs.Ultimate_SlowDown;
       #Ultimate_Creep := #VTD_Control.Inputs.Ultimate_Creep;
       #Lower_Limit := #VTD_Control.Inputs.Lower_Limit;
       #Level_Detect1 := #VTD_Control.Inputs.Level_Detect1;
       #Level_Detect2 := #VTD_Control.Inputs.Level_Detect2;
       #DP1_Extended := #VTD_Control.Inputs.DP1_Extended;
       #DP1_Retracted := #VTD_Control.Inputs.DP1_Retracted;
       #DP2_Extended := #VTD_Control.Inputs.DP2_Extended;
       #DP2_Retracted := #VTD_Control.Inputs.DP2_Retracted;
       #Chain_Slack_1 := #VTD_Control.Inputs.Chain_Slack_1;
       #Chain_Slack_2 := #VTD_Control.Inputs.Chain_Slack_2;
       #Chain_Slack_3 := #VTD_Control.Inputs.Chain_Slack_3;
       #Chain_Slack_4 := #VTD_Control.Inputs.Chain_Slack_4;
       #Shuttle_Detect1 := #Cnv_Sensors.Overhang_Left;
       #Shuttle_Detect2 := #Cnv_Sensors.Overhang_Right;
       #VTD_Control.LE := #VTD_Control.Inputs.LE_Position;
       #VTD_Control.AE := #VTD_Control.Inputs.AE_Position_1;
   END_REGION

   REGION Cyclic Checks
       // Check for shuttle
       IF #System_no > 3 THEN
           IF #Shuttle_Detect1 AND #Shuttle_Detect2 THEN
               #VTD_Control.Shuttle_Loaded := 1; //inplace
           ELSIF NOT #Shuttle_Detect1 AND #Shuttle_Detect2 THEN
               #VTD_Control.Shuttle_Loaded := 2; // Front overhang
           ELSIF #Shuttle_Detect1 AND NOT #Shuttle_Detect2 THEN
               #VTD_Control.Shuttle_Loaded := 3; //Rear overhang
           ELSE
               #VTD_Control.Shuttle_Loaded := 0; //None
           END_IF;
       END_IF;

       // Check for Pallet
       IF #Cnv_Sensors.Left OR #Cnv_Sensors.Lpd1 OR #Cnv_Sensors.Center OR #Cnv_Sensors.Rpd1 OR #Cnv_Sensors.Right THEN
           //Chep Pallet
           IF #Cnv_Sensors.Left AND #Cnv_Sensors.Right THEN
               #VTD_Control.Pallet_Loaded := #CHEP;//Chep
               //Euro skewed to the left (BACK)
           ELSIF #Cnv_Sensors.Rpd1 AND #Cnv_Sensors.Left AND NOT #Cnv_Sensors.Right THEN
               #VTD_Control.Pallet_Loaded := #"EURO LEFT";//'Euro BACK';
               //Euro skewed to the right (FRONT)
           ELSIF #Cnv_Sensors.Lpd1 AND #Cnv_Sensors.Right AND NOT #Cnv_Sensors.Left THEN
               #VTD_Control.Pallet_Loaded := #"EURO RIGHT";//'Euro FRONT';
               //Euro CENTERED
           ELSIF #Cnv_Sensors.Center AND #Cnv_Sensors.Lpd1 AND #Cnv_Sensors.Rpd1 THEN
               #VTD_Control.Pallet_Loaded := #"EURO CENTER";//'Euro centered';
               //Some unknown combination of Cnv_Inputs
           ELSE
               #VTD_Control.Pallet_Loaded := #UNKNOWN;//'Unknown';
           END_IF;
       ELSE
           //No Pallet
           #VTD_Control.Pallet_Loaded := #EMPTY;//'None';
       END_IF;

       //Docking pins
           IF #DP1_Extended AND #DP2_Extended THEN
               #VTD_Control.LP_State := 1; //'Extended'
           ELSIF #DP1_Retracted AND #DP2_Retracted THEN
               #VTD_Control.LP_State := 2; //'Retracted'
           ELSE
               #VTD_Control.LP_State := 0; //'Unknown'
           END_IF;

           #VTD_Control.DP_Extended := #VTD_Control.LP_State = 1;

       // Level detect
       #Level_Detect := #Level_Detect1 AND #Level_Detect2;

       //VTD extractor is docked
       IF #DP1_Extended AND #DP2_Extended AND #Level_Detect AND
           (#VTD_Control.LE - #VTD_Settings.Teach_Values.Levels_LE[#LevelBelowExtractor]) <= #VTD_Settings.Level_Detect_LE THEN
           #VTD_Control.Docked := TRUE;
       ELSE
           #VTD_Control.Docked := FALSE;
       END_IF;

       //Ultimate stop checks
       IF (#VTD_Control.LE < #VTD_Settings.Slowdown_Count_LE OR #VTD_Control.LE > #VTD_Settings.Teach_Values.Levels_LE[#VTD_Settings.Highest_Level] - #VTD_Settings.Slowdown_Count_LE) AND
           #Ultimate_Creep AND #Ultimate_SlowDown AND #VTD_Control.Running THEN
           #VTD_Control.Motor_Speed := #VTD_Settings.Creep_Speed;
           #VTD_Control.Warning := 3; // Overtravel creep zone reached
       ELSIF (#VTD_Control.LE < #VTD_Settings.Slowdown_Count_LE OR #VTD_Control.LE > #VTD_Settings.Teach_Values.Levels_LE[#VTD_Settings.Highest_Level] - #VTD_Settings.Slowdown_Count_LE) AND
           NOT #Ultimate_Creep AND #Ultimate_SlowDown AND #VTD_Control.Running THEN
           #VTD_Control.Motor_Speed := #VTD_Settings.Slow_Speed; // Overtravel slow zone reached
       END_IF;

       //Update Variables
       IF #VTD_Control.Current_Task_Type = 0 OR #VTD_Control.Current_Task_Type = 1 THEN
           #VTD_Control.SM_State := #State;
       ELSIF #VTD_Control.Current_Task_Type = 2 OR #VTD_Control.Current_Task_Type = 3 THEN
           #VTD_Control.SM_State := #I_State;
       END_IF;

       FOR #i := #VTD_Settings.Lowest_Level TO #VTD_Settings.Highest_Level DO
           IF NOT "Control_DB".LCnv_Sys[#System_no].Cnv_Level[#i].Cnv1.Safety_Stop_Cnrl.Inputs.DP_Extended THEN
               #Cnvs1_NotExtended := true;
           END_IF;
           IF NOT "Control_DB".LCnv_Sys[#System_no].Cnv_Level[#i].Cnv2.Safety_Stop_Cnrl.Inputs.DP_Extended THEN
               #Cnvs2_NotExtended := true;
           END_IF;
       END_FOR;

       //Confirm whish level is below the extractor
       FOR #i := #VTD_Settings.Lowest_Level TO #VTD_Settings.Highest_Level DO
           IF #VTD_Control.LE >= (#VTD_Settings.Teach_Values.Levels_LE[#i] - #VTD_Settings.Level_Detect_LE) THEN
               #LevelBelowExtractor := #i;
           END_IF;
       END_FOR;

       #Stoppers_NotExtended := #Cnvs1_NotExtended (*AND #Cnvs2_NotExtended*);

       //AE ERROR
       IF #VTD_Control.Inputs.AE_Status_2.%X15 THEN
           #VTD_Control.AE_Error := 1;
       ELSE
           #VTD_Control.AE_Error := 0;
       END_IF;

       //Encoder Delta
       #VTD_Control.Encoder_Delta := ABS(#VTD_Control.AE - #VTD_Control.LE);

       //CURRENT LEVEL
       FOR #i := #VTD_Settings.Lowest_Level TO #VTD_Settings.Highest_Level DO
           IF ABS(#VTD_Control.LE - #VTD_Settings.Teach_Values.Levels_LE[#i]) <= #VTD_Settings.VTD_Level_Granularity AND #Level_Detect THEN
               #VTD_Control.Current_Level := #i;
               EXIT;
           ELSE
               #VTD_Control.Current_Level := 0;
           END_IF;
       END_FOR;

       //SPEED mm/S
       #T_Speed(IN := TRUE,
                PT := T#100MS);

       IF #T_Speed.Q THEN
           #DeltaPos_mm := ABS(#VTD_Control.LE - #LE_Prev_mm);
           #VTDSpeed_mm_s := #DeltaPos_mm / #SampleTime_s;
           #LE_Prev_mm := #VTD_Control.LE;
           #T_Speed(IN := FALSE,
                    PT := T#0MS);
       END_IF;
   END_REGION

   REGION Auto/Semi-Auto Mode
       CASE #State OF
           0: //Idle
               #Last_State := #State;
               #VTD_Control.Motor_UP := FALSE;
               #VTD_Control.Motor_Down := FALSE;
               #VTD_Control.Motor.Speed := 0;
               #DestinationLevel := #CurrentlLevel := 0;
               #VTD_Control.Stopped := TRUE;
               #Watchdog.TON(IN := FALSE,
                             PT := T#0S);
               IF #VTD_Control.Mode = 3 OR #VTD_Control.Mode = 2 THEN
                   IF #VTD_Control.Instruction.Enable AND NOT #VTD_Control.Error THEN
                       #State := 10;
                   END_IF;
               END_IF;

           10: //Standby
               #Last_State := #State;
               IF #VTD_Control.Enabled AND NOT #VTD_Control.Running AND #VTD_Control.Instruction.Move_To_Level >= #VTD_Settings.Lowest_Level AND
                   #VTD_Control.Instruction.Move_To_Level <= #VTD_Settings.Highest_Level AND #VTD_Control.Pallet_Loaded <> #UNKNOWN AND
                   ((#VTD_Control.Instruction.Task_ID > 0 OR #VTD_Control.Instruction.Task_Metadata <> '' AND #VTD_Control.Mode = 3 AND "Control_DB".WCS_OPC_Control[#System_no].Task_Type = 1) OR
                   (#VTD_Control.Mode = 2 (*AND #R_Execulte.Q*)))
               THEN
                   IF (#VTD_Control.Instruction.Move_To_Level = #VTD_Control.Current_Level AND #VTD_Control.Instruction.Move_To_Level <> 0) OR "Control_DB".ECnv_Sys[#System_no].Running THEN
                       #VTD_Control.Warning := 1; //VTD already at level requested
                       #VTD_Control.Instruction.Move_To_Level := 0;
                       //Go straght to the travel complete feedabck 
                   ELSIF #VTD_Control.Shuttle_Loaded = 0 OR #VTD_Control.Shuttle_Loaded = 1
                   THEN //EVERYTHING OK
                       #DestinationLevel := #VTD_Control.Instruction.Move_To_Level;
                       #CurrentlLevel := #VTD_Control.Current_Level;
                       #VTD_Control.Current_Task_ID := #VTD_Control.Instruction.Task_ID;
                       #VTD_Control.Running := TRUE;
                       #State := 20;
                   END_IF;
               END_IF;

           20: //Extend all safety stoppers that are not in the up position
               #Last_State := #State;
               #VTD_Control.Done := FALSE;// To report to order table
               FOR #i := #VTD_Settings.Lowest_Level TO #VTD_Settings.Highest_Level DO
                   IF NOT "Control_DB".LCnv_Sys[#System_no].Cnv_Level[#i].Cnv1.Safety_Stop_Cnrl.Inputs.DP_Extended THEN
                       "Control_DB".LCnv_Sys[#System_no].Cnv_Level[#i].Cnv1.Safety_Stop_Cnrl.Instruction.Extend := TRUE;
                   END_IF;
                   IF NOT "Control_DB".LCnv_Sys[#System_no].Cnv_Level[#i].Cnv2.Safety_Stop_Cnrl.Inputs.DP_Extended THEN
                       "Control_DB".LCnv_Sys[#System_no].Cnv_Level[#i].Cnv2.Safety_Stop_Cnrl.Instruction.Extend := TRUE;
                   END_IF;
               END_FOR;
               #State := 25;

           25: //Check to ensure the Safety stoppers are in the up position.
               #Last_State := #State;
               FOR #i := #VTD_Settings.Lowest_Level TO #VTD_Settings.Highest_Level DO
                   IF "Control_DB".LCnv_Sys[#System_no].Cnv_Level[#i].Cnv1.Safety_Stop_Cnrl.Inputs.DP_Extended THEN
                       "Control_DB".LCnv_Sys[#System_no].Cnv_Level[#i].Cnv1.Safety_Stop_Cnrl.Instruction.Extend := FALSE;
                   END_IF;
                   IF "Control_DB".LCnv_Sys[#System_no].Cnv_Level[#i].Cnv2.Safety_Stop_Cnrl.Inputs.DP_Extended THEN
                       "Control_DB".LCnv_Sys[#System_no].Cnv_Level[#i].Cnv2.Safety_Stop_Cnrl.Instruction.Extend := FALSE;
                   END_IF;
               END_FOR;
               IF  ("Control_DB".LCnv_Sys[#System_no].Cnv_Level[1].Cnv1.Safety_Stop_Cnrl.Inputs.DP_Extended OR #System_no <= 3) AND
                   "Control_DB".LCnv_Sys[#System_no].Cnv_Level[2].Cnv1.Safety_Stop_Cnrl.Inputs.DP_Extended AND
                   "Control_DB".LCnv_Sys[#System_no].Cnv_Level[3].Cnv1.Safety_Stop_Cnrl.Inputs.DP_Extended AND
                   "Control_DB".LCnv_Sys[#System_no].Cnv_Level[4].Cnv1.Safety_Stop_Cnrl.Inputs.DP_Extended AND
                   "Control_DB".LCnv_Sys[#System_no].Cnv_Level[5].Cnv1.Safety_Stop_Cnrl.Inputs.DP_Extended AND
                   "Control_DB".LCnv_Sys[#System_no].Cnv_Level[6].Cnv1.Safety_Stop_Cnrl.Inputs.DP_Extended AND
                   "Control_DB".LCnv_Sys[#System_no].Cnv_Level[7].Cnv1.Safety_Stop_Cnrl.Inputs.DP_Extended AND
                   "Control_DB".LCnv_Sys[#System_no].Cnv_Level[8].Cnv1.Safety_Stop_Cnrl.Inputs.DP_Extended AND
                   "Control_DB".LCnv_Sys[#System_no].Cnv_Level[2].Cnv2.Safety_Stop_Cnrl.Inputs.DP_Extended AND
                   "Control_DB".LCnv_Sys[#System_no].Cnv_Level[3].Cnv2.Safety_Stop_Cnrl.Inputs.DP_Extended AND
                   "Control_DB".LCnv_Sys[#System_no].Cnv_Level[4].Cnv2.Safety_Stop_Cnrl.Inputs.DP_Extended AND
                   "Control_DB".LCnv_Sys[#System_no].Cnv_Level[5].Cnv2.Safety_Stop_Cnrl.Inputs.DP_Extended AND
                   "Control_DB".LCnv_Sys[#System_no].Cnv_Level[6].Cnv2.Safety_Stop_Cnrl.Inputs.DP_Extended AND
                   "Control_DB".LCnv_Sys[#System_no].Cnv_Level[7].Cnv2.Safety_Stop_Cnrl.Inputs.DP_Extended AND
                   "Control_DB".LCnv_Sys[#System_no].Cnv_Level[8].Cnv2.Safety_Stop_Cnrl.Inputs.DP_Extended
               THEN
                   #State := 30;
                   #Stopper_Extend_Timer(IN := FALSE,PT := T#0s); // Reset the timer, safety stoppers up
               ELSE
                   #Stopper_Extend_Timer(IN := TRUE,
                                         PT := UINT_TO_TIME("Settings_DB".LCnv_Sys[#System_no].Cnv_Level[2].Cnv1.Safety_stop_Timeout)); // ascent time 
                   IF #Stopper_Extend_Timer.Q THEN
                       "Set_Bit_F"(Bit := 6, // safety stopper error during VTD sequence
                                   Bit_Value := 1,
                                   Var := #VTD_Control.VTD_Errors.Error_Word_2);

